Yaskawa INFORM job: ITEST.JBI

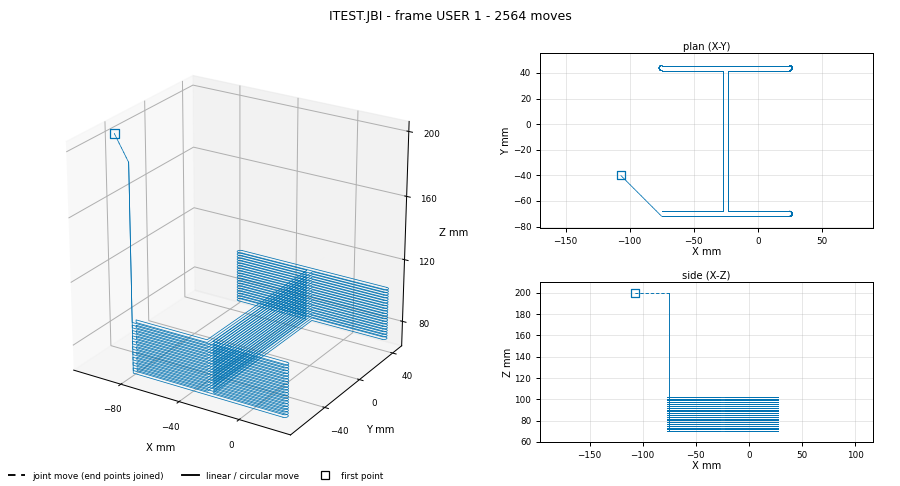
[picture p0: tool path of ITEST.JBI in frame USER 1, 2564 of 2624 moves have a stored position in this frame; points joined in program order, loops and branches not executed]
/JOB
//NAME ITEST
//POS
///NPOS 2624,0,0,0,0,0
///USER 1
///TOOL 1
///POSTYPE USER
///RECTAN
///RCONF 1,0,0,0,0,0,0,0,0,0,0,0,0,0,0,0,0,0,0,0,0,0,0,0
C00000=-107.000,-40.000,200.000,0.0000,0.0000,-150.0000
C00001=-75.000,-72.000,200.000,0.0000,0.0000,-150.0000
C00002=-75.000,-72.000,70.000,0.0000,0.0000,-150.0000
C00003=-70.000,-72.000,70.000,0.0000,0.0000,-150.0000
C00004=-65.000,-72.000,70.000,0.0000,0.0000,-150.0000
C00005=-60.000,-72.000,70.000,0.0000,0.0000,-150.0000
C00006=-55.000,-72.000,70.000,0.0000,0.0000,-150.0000
C00007=-50.000,-72.000,70.000,0.0000,0.0000,-150.0000
C00008=-45.000,-72.000,70.000,0.0000,0.0000,-150.0000
C00009=-40.000,-72.000,70.000,0.0000,0.0000,-150.0000
C00010=-35.000,-72.000,70.000,0.0000,0.0000,-150.0000
C00011=-30.000,-72.000,70.000,0.0000,0.0000,-150.0000
C00012=-25.000,-72.000,70.000,0.0000,0.0000,-150.0000
C00013=-20.000,-72.000,70.000,0.0000,0.0000,-150.0000
C00014=-15.000,-72.000,70.000,0.0000,0.0000,-150.0000
C00015=-10.000,-72.000,70.000,0.0000,0.0000,-150.0000
C00016=-5.000,-72.000,70.000,0.0000,0.0000,-150.0000
C00017=0.000,-72.000,70.000,0.0000,0.0000,-150.0000
C00018=5.000,-72.000,70.000,0.0000,0.0000,-150.0000
C00019=10.000,-72.000,70.000,0.0000,0.0000,-150.0000
C00020=15.000,-72.000,70.000,0.0000,0.0000,-150.0000
C00021=20.000,-72.000,70.000,0.0000,0.0000,-150.0000
C00022=25.000,-72.000,70.000,0.0000,0.0000,-150.0000
C00023=26.950,-70.050,70.000,0.0000,0.0000,-150.0000
C00024=25.000,-68.100,70.000,0.0000,0.0000,-150.0000
C00025=20.195,-68.100,70.000,0.0000,0.0000,-150.0000
C00026=15.390,-68.100,70.000,0.0000,0.0000,-150.0000
C00027=10.585,-68.100,70.000,0.0000,0.0000,-150.0000
C00028=5.780,-68.100,70.000,0.0000,0.0000,-150.0000
C00029=0.975,-68.100,70.000,0.0000,0.0000,-150.0000
C00030=-3.830,-68.100,70.000,0.0000,0.0000,-150.0000
C00031=-8.635,-68.100,70.000,0.0000,0.0000,-150.0000
C00032=-13.440,-68.100,70.000,0.0000,0.0000,-150.0000
C00033=-18.245,-68.100,70.000,0.0000,0.0000,-150.0000
C00034=-23.050,-68.100,70.000,0.0000,0.0000,-150.0000
C00035=-23.050,-63.100,70.000,0.0000,0.0000,-150.0000
C00036=-23.050,-58.100,70.000,0.0000,0.0000,-150.0000
C00037=-23.050,-53.100,70.000,0.0000,0.0000,-150.0000
C00038=-23.050,-48.100,70.000,0.0000,0.0000,-150.0000
C00039=-23.050,-43.100,70.000,0.0000,0.0000,-150.0000
C00040=-23.050,-38.100,70.000,0.0000,0.0000,-150.0000
C00041=-23.050,-33.100,70.000,0.0000,0.0000,-150.0000
C00042=-23.050,-28.100,70.000,0.0000,0.0000,-150.0000
C00043=-23.050,-23.100,70.000,0.0000,0.0000,-150.0000
C00044=-23.050,-18.100,70.000,0.0000,0.0000,-150.0000
C00045=-23.050,-13.100,70.000,0.0000,0.0000,-150.0000
C00046=-23.050,-8.100,70.000,0.0000,0.0000,-150.0000
C00047=-23.050,-3.100,70.000,0.0000,0.0000,-150.0000
C00048=-23.050,1.900,70.000,0.0000,0.0000,-150.0000
C00049=-23.050,6.900,70.000,0.0000,0.0000,-150.0000
C00050=-23.050,11.900,70.000,0.0000,0.0000,-150.0000
C00051=-23.050,16.900,70.000,0.0000,0.0000,-150.0000
C00052=-23.050,21.900,70.000,0.0000,0.0000,-150.0000
C00053=-23.050,26.900,70.000,0.0000,0.0000,-150.0000
C00054=-23.050,31.900,70.000,0.0000,0.0000,-150.0000
C00055=-23.050,36.900,70.000,0.0000,0.0000,-150.0000
C00056=-23.050,41.900,70.000,0.0000,0.0000,-150.0000
C00057=-18.267,41.900,70.000,0.0000,0.0000,-150.0000
C00058=-13.483,41.900,70.000,0.0000,0.0000,-150.0000
C00059=-8.700,41.900,70.000,0.0000,0.0000,-150.0000
C00060=-3.917,41.900,70.000,0.0000,0.0000,-150.0000
C00061=0.867,41.900,70.000,0.0000,0.0000,-150.0000
C00062=5.650,41.900,70.000,0.0000,0.0000,-150.0000
C00063=10.433,41.900,70.000,0.0000,0.0000,-150.0000
C00064=15.217,41.900,70.000,0.0000,0.0000,-150.0000
C00065=20.000,41.900,70.000,0.0000,0.0000,-150.0000
C00066=25.000,41.900,70.000,0.0000,0.0000,-150.0000
C00067=26.950,43.850,70.000,0.0000,0.0000,-150.0000
C00068=25.000,45.800,70.000,0.0000,0.0000,-150.0000
C00069=20.000,45.800,70.000,0.0000,0.0000,-150.0000
C00070=15.000,45.800,70.000,0.0000,0.0000,-150.0000
C00071=10.000,45.800,70.000,0.0000,0.0000,-150.0000
C00072=5.000,45.800,70.000,0.0000,0.0000,-150.0000
C00073=0.000,45.800,70.000,0.0000,0.0000,-150.0000
C00074=-5.000,45.800,70.000,0.0000,0.0000,-150.0000
C00075=-10.000,45.800,70.000,0.0000,0.0000,-150.0000
C00076=-15.000,45.800,70.000,0.0000,0.0000,-150.0000
C00077=-20.000,45.800,70.000,0.0000,0.0000,-150.0000
C00078=-25.000,45.800,70.000,0.0000,0.0000,-150.0000
C00079=-30.000,45.800,70.000,0.0000,0.0000,-150.0000
C00080=-35.000,45.800,70.000,0.0000,0.0000,-150.0000
C00081=-40.000,45.800,70.000,0.0000,0.0000,-150.0000
C00082=-45.000,45.800,70.000,0.0000,0.0000,-150.0000
C00083=-50.000,45.800,70.000,0.0000,0.0000,-150.0000
C00084=-55.000,45.800,70.000,0.0000,0.0000,-150.0000
C00085=-60.000,45.800,70.000,0.0000,0.0000,-150.0000
C00086=-65.000,45.800,70.000,0.0000,0.0000,-150.0000
C00087=-70.000,45.800,70.000,0.0000,0.0000,-150.0000
C00088=-75.000,45.800,70.000,0.0000,0.0000,-150.0000
C00089=-76.950,43.850,70.000,0.0000,0.0000,-150.0000
C00090=-75.000,41.900,70.000,0.0000,0.0000,-150.0000
C00091=-70.195,41.900,70.000,0.0000,0.0000,-150.0000
C00092=-65.390,41.900,70.000,0.0000,0.0000,-150.0000
C00093=-60.585,41.900,70.000,0.0000,0.0000,-150.0000
C00094=-55.780,41.900,70.000,0.0000,0.0000,-150.0000
C00095=-50.975,41.900,70.000,0.0000,0.0000,-150.0000
C00096=-46.170,41.900,70.000,0.0000,0.0000,-150.0000
C00097=-41.365,41.900,70.000,0.0000,0.0000,-150.0000
C00098=-36.560,41.900,70.000,0.0000,0.0000,-150.0000
C00099=-31.755,41.900,70.000,0.0000,0.0000,-150.0000
C00100=-26.950,41.900,70.000,0.0000,0.0000,-150.0000
C00101=-26.950,36.900,70.000,0.0000,0.0000,-150.0000
C00102=-26.950,31.900,70.000,0.0000,0.0000,-150.0000
C00103=-26.950,26.900,70.000,0.0000,0.0000,-150.0000
C00104=-26.950,21.900,70.000,0.0000,0.0000,-150.0000
C00105=-26.950,16.900,70.000,0.0000,0.0000,-150.0000
C00106=-26.950,11.900,70.000,0.0000,0.0000,-150.0000
C00107=-26.950,6.900,70.000,0.0000,0.0000,-150.0000
C00108=-26.950,1.900,70.000,0.0000,0.0000,-150.0000
C00109=-26.950,-3.100,70.000,0.0000,0.0000,-150.0000
C00110=-26.950,-8.100,70.000,0.0000,0.0000,-150.0000
C00111=-26.950,-13.100,70.000,0.0000,0.0000,-150.0000
C00112=-26.950,-18.100,70.000,0.0000,0.0000,-150.0000
C00113=-26.950,-23.100,70.000,0.0000,0.0000,-150.0000
C00114=-26.950,-28.100,70.000,0.0000,0.0000,-150.0000
C00115=-26.950,-33.100,70.000,0.0000,0.0000,-150.0000
C00116=-26.950,-38.100,70.000,0.0000,0.0000,-150.0000
C00117=-26.950,-43.100,70.000,0.0000,0.0000,-150.0000
C00118=-26.950,-48.100,70.000,0.0000,0.0000,-150.0000
C00119=-26.950,-53.100,70.000,0.0000,0.0000,-150.0000
C00120=-26.950,-58.100,70.000,0.0000,0.0000,-150.0000
C00121=-26.950,-63.100,70.000,0.0000,0.0000,-150.0000
C00122=-26.950,-68.100,70.000,0.0000,0.0000,-150.0000
C00123=-31.755,-68.100,70.000,0.0000,0.0000,-150.0000
C00124=-36.560,-68.100,70.000,0.0000,0.0000,-150.0000
C00125=-41.365,-68.100,70.000,0.0000,0.0000,-150.0000
C00126=-46.170,-68.100,70.000,0.0000,0.0000,-150.0000
C00127=-50.975,-68.100,70.000,0.0000,0.0000,-150.0000
C00128=-55.780,-68.100,70.000,0.0000,0.0000,-150.0000
C00129=-60.585,-68.100,70.000,0.0000,0.0000,-150.0000
C00130=-65.390,-68.100,70.000,0.0000,0.0000,-150.0000
C00131=-70.195,-68.100,70.000,0.0000,0.0000,-150.0000
C00132=-75.000,-68.100,70.000,0.0000,0.0000,-150.0000
C00133=-75.000,-68.100,71.700,0.0000,0.0000,-150.0000
C00134=-70.195,-68.100,71.700,0.0000,0.0000,-150.0000
C00135=-65.390,-68.100,71.700,0.0000,0.0000,-150.0000
C00136=-60.585,-68.100,71.700,0.0000,0.0000,-150.0000
C00137=-55.780,-68.100,71.700,0.0000,0.0000,-150.0000
C00138=-50.975,-68.100,71.700,0.0000,0.0000,-150.0000
C00139=-46.170,-68.100,71.700,0.0000,0.0000,-150.0000
C00140=-41.365,-68.100,71.700,0.0000,0.0000,-150.0000
C00141=-36.560,-68.100,71.700,0.0000,0.0000,-150.0000
C00142=-31.755,-68.100,71.700,0.0000,0.0000,-150.0000
C00143=-26.950,-68.100,71.700,0.0000,0.0000,-150.0000
C00144=-26.950,-63.100,71.700,0.0000,0.0000,-150.0000
C00145=-26.950,-58.100,71.700,0.0000,0.0000,-150.0000
C00146=-26.950,-53.100,71.700,0.0000,0.0000,-150.0000
C00147=-26.950,-48.100,71.700,0.0000,0.0000,-150.0000
C00148=-26.950,-43.100,71.700,0.0000,0.0000,-150.0000
C00149=-26.950,-38.100,71.700,0.0000,0.0000,-150.0000
C00150=-26.950,-33.100,71.700,0.0000,0.0000,-150.0000
C00151=-26.950,-28.100,71.700,0.0000,0.0000,-150.0000
C00152=-26.950,-23.100,71.700,0.0000,0.0000,-150.0000
C00153=-26.950,-18.100,71.700,0.0000,0.0000,-150.0000
C00154=-26.950,-13.100,71.700,0.0000,0.0000,-150.0000
C00155=-26.950,-8.100,71.700,0.0000,0.0000,-150.0000
C00156=-26.950,-3.100,71.700,0.0000,0.0000,-150.0000
C00157=-26.950,1.900,71.700,0.0000,0.0000,-150.0000
C00158=-26.950,6.900,71.700,0.0000,0.0000,-150.0000
C00159=-26.950,11.900,71.700,0.0000,0.0000,-150.0000
C00160=-26.950,16.900,71.700,0.0000,0.0000,-150.0000
C00161=-26.950,21.900,71.700,0.0000,0.0000,-150.0000
C00162=-26.950,26.900,71.700,0.0000,0.0000,-150.0000
C00163=-26.950,31.900,71.700,0.0000,0.0000,-150.0000
C00164=-26.950,36.900,71.700,0.0000,0.0000,-150.0000
C00165=-26.950,41.900,71.700,0.0000,0.0000,-150.0000
C00166=-31.733,41.900,71.700,0.0000,0.0000,-150.0000
C00167=-36.517,41.900,71.700,0.0000,0.0000,-150.0000
C00168=-41.300,41.900,71.700,0.0000,0.0000,-150.0000
C00169=-46.083,41.900,71.700,0.0000,0.0000,-150.0000
C00170=-50.867,41.900,71.700,0.0000,0.0000,-150.0000
C00171=-55.650,41.900,71.700,0.0000,0.0000,-150.0000
C00172=-60.433,41.900,71.700,0.0000,0.0000,-150.0000
C00173=-65.217,41.900,71.700,0.0000,0.0000,-150.0000
C00174=-70.000,41.900,71.700,0.0000,0.0000,-150.0000
C00175=-75.000,41.900,71.700,0.0000,0.0000,-150.0000
C00176=-76.950,43.850,71.700,0.0000,0.0000,-150.0000
C00177=-75.000,45.800,71.700,0.0000,0.0000,-150.0000
C00178=-70.000,45.800,71.700,0.0000,0.0000,-150.0000
C00179=-65.000,45.800,71.700,0.0000,0.0000,-150.0000
C00180=-60.000,45.800,71.700,0.0000,0.0000,-150.0000
C00181=-55.000,45.800,71.700,0.0000,0.0000,-150.0000
C00182=-50.000,45.800,71.700,0.0000,0.0000,-150.0000
C00183=-45.000,45.800,71.700,0.0000,0.0000,-150.0000
C00184=-40.000,45.800,71.700,0.0000,0.0000,-150.0000
C00185=-35.000,45.800,71.700,0.0000,0.0000,-150.0000
C00186=-30.000,45.800,71.700,0.0000,0.0000,-150.0000
C00187=-25.000,45.800,71.700,0.0000,0.0000,-150.0000
C00188=-20.000,45.800,71.700,0.0000,0.0000,-150.0000
C00189=-15.000,45.800,71.700,0.0000,0.0000,-150.0000
C00190=-10.000,45.800,71.700,0.0000,0.0000,-150.0000
C00191=-5.000,45.800,71.700,0.0000,0.0000,-150.0000
C00192=0.000,45.800,71.700,0.0000,0.0000,-150.0000
C00193=5.000,45.800,71.700,0.0000,0.0000,-150.0000
C00194=10.000,45.800,71.700,0.0000,0.0000,-150.0000
C00195=15.000,45.800,71.700,0.0000,0.0000,-150.0000
C00196=20.000,45.800,71.700,0.0000,0.0000,-150.0000
C00197=25.000,45.800,71.700,0.0000,0.0000,-150.0000
C00198=26.950,43.850,71.700,0.0000,0.0000,-150.0000
C00199=25.000,41.900,71.700,0.0000,0.0000,-150.0000
C00200=20.195,41.900,71.700,0.0000,0.0000,-150.0000
C00201=15.390,41.900,71.700,0.0000,0.0000,-150.0000
C00202=10.585,41.900,71.700,0.0000,0.0000,-150.0000
C00203=5.780,41.900,71.700,0.0000,0.0000,-150.0000
C00204=0.975,41.900,71.700,0.0000,0.0000,-150.0000
C00205=-3.830,41.900,71.700,0.0000,0.0000,-150.0000
C00206=-8.635,41.900,71.700,0.0000,0.0000,-150.0000
C00207=-13.440,41.900,71.700,0.0000,0.0000,-150.0000
C00208=-18.245,41.900,71.700,0.0000,0.0000,-150.0000
C00209=-23.050,41.900,71.700,0.0000,0.0000,-150.0000
C00210=-23.050,36.900,71.700,0.0000,0.0000,-150.0000
C00211=-23.050,31.900,71.700,0.0000,0.0000,-150.0000
C00212=-23.050,26.900,71.700,0.0000,0.0000,-150.0000
C00213=-23.050,21.900,71.700,0.0000,0.0000,-150.0000
C00214=-23.050,16.900,71.700,0.0000,0.0000,-150.0000
C00215=-23.050,11.900,71.700,0.0000,0.0000,-150.0000
C00216=-23.050,6.900,71.700,0.0000,0.0000,-150.0000
C00217=-23.050,1.900,71.700,0.0000,0.0000,-150.0000
C00218=-23.050,-3.100,71.700,0.0000,0.0000,-150.0000
C00219=-23.050,-8.100,71.700,0.0000,0.0000,-150.0000
C00220=-23.050,-13.100,71.700,0.0000,0.0000,-150.0000
C00221=-23.050,-18.100,71.700,0.0000,0.0000,-150.0000
C00222=-23.050,-23.100,71.700,0.0000,0.0000,-150.0000
C00223=-23.050,-28.100,71.700,0.0000,0.0000,-150.0000
C00224=-23.050,-33.100,71.700,0.0000,0.0000,-150.0000
C00225=-23.050,-38.100,71.700,0.0000,0.0000,-150.0000
C00226=-23.050,-43.100,71.700,0.0000,0.0000,-150.0000
C00227=-23.050,-48.100,71.700,0.0000,0.0000,-150.0000
C00228=-23.050,-53.100,71.700,0.0000,0.0000,-150.0000
C00229=-23.050,-58.100,71.700,0.0000,0.0000,-150.0000
C00230=-23.050,-63.100,71.700,0.0000,0.0000,-150.0000
C00231=-23.050,-68.100,71.700,0.0000,0.0000,-150.0000
C00232=-18.267,-68.100,71.700,0.0000,0.0000,-150.0000
C00233=-13.483,-68.100,71.700,0.0000,0.0000,-150.0000
C00234=-8.700,-68.100,71.700,0.0000,0.0000,-150.0000
C00235=-3.917,-68.100,71.700,0.0000,0.0000,-150.0000
C00236=0.867,-68.100,71.700,0.0000,0.0000,-150.0000
C00237=5.650,-68.100,71.700,0.0000,0.0000,-150.0000
C00238=10.433,-68.100,71.700,0.0000,0.0000,-150.0000
C00239=15.217,-68.100,71.700,0.0000,0.0000,-150.0000
C00240=20.000,-68.100,71.700,0.0000,0.0000,-150.0000
C00241=25.000,-68.100,71.700,0.0000,0.0000,-150.0000
C00242=26.950,-70.050,71.700,0.0000,0.0000,-150.0000
C00243=25.000,-72.000,71.700,0.0000,0.0000,-150.0000
C00244=20.000,-72.000,71.700,0.0000,0.0000,-150.0000
C00245=15.000,-72.000,71.700,0.0000,0.0000,-150.0000
C00246=10.000,-72.000,71.700,0.0000,0.0000,-150.0000
C00247=5.000,-72.000,71.700,0.0000,0.0000,-150.0000
C00248=0.000,-72.000,71.700,0.0000,0.0000,-150.0000
C00249=-5.000,-72.000,71.700,0.0000,0.0000,-150.0000
C00250=-10.000,-72.000,71.700,0.0000,0.0000,-150.0000
C00251=-15.000,-72.000,71.700,0.0000,0.0000,-150.0000
C00252=-20.000,-72.000,71.700,0.0000,0.0000,-150.0000
C00253=-25.000,-72.000,71.700,0.0000,0.0000,-150.0000
C00254=-30.000,-72.000,71.700,0.0000,0.0000,-150.0000
C00255=-35.000,-72.000,71.700,0.0000,0.0000,-150.0000
C00256=-40.000,-72.000,71.700,0.0000,0.0000,-150.0000
C00257=-45.000,-72.000,71.700,0.0000,0.0000,-150.0000
C00258=-50.000,-72.000,71.700,0.0000,0.0000,-150.0000
C00259=-55.000,-72.000,71.700,0.0000,0.0000,-150.0000
C00260=-60.000,-72.000,71.700,0.0000,0.0000,-150.0000
C00261=-65.000,-72.000,71.700,0.0000,0.0000,-150.0000
C00262=-70.000,-72.000,71.700,0.0000,0.0000,-150.0000
C00263=-75.000,-72.000,71.700,0.0000,0.0000,-150.0000
C00264=-75.000,-72.000,73.400,0.0000,0.0000,-150.0000
C00265=-70.000,-72.000,73.400,0.0000,0.0000,-150.0000
C00266=-65.000,-72.000,73.400,0.0000,0.0000,-150.0000
C00267=-60.000,-72.000,73.400,0.0000,0.0000,-150.0000
C00268=-55.000,-72.000,73.400,0.0000,0.0000,-150.0000
C00269=-50.000,-72.000,73.400,0.0000,0.0000,-150.0000
C00270=-45.000,-72.000,73.400,0.0000,0.0000,-150.0000
C00271=-40.000,-72.000,73.400,0.0000,0.0000,-150.0000
C00272=-35.000,-72.000,73.400,0.0000,0.0000,-150.0000
C00273=-30.000,-72.000,73.400,0.0000,0.0000,-150.0000
C00274=-25.000,-72.000,73.400,0.0000,0.0000,-150.0000
C00275=-20.000,-72.000,73.400,0.0000,0.0000,-150.0000
C00276=-15.000,-72.000,73.400,0.0000,0.0000,-150.0000
C00277=-10.000,-72.000,73.400,0.0000,0.0000,-150.0000
C00278=-5.000,-72.000,73.400,0.0000,0.0000,-150.0000
C00279=0.000,-72.000,73.400,0.0000,0.0000,-150.0000
C00280=5.000,-72.000,73.400,0.0000,0.0000,-150.0000
C00281=10.000,-72.000,73.400,0.0000,0.0000,-150.0000
C00282=15.000,-72.000,73.400,0.0000,0.0000,-150.0000
C00283=20.000,-72.000,73.400,0.0000,0.0000,-150.0000
C00284=25.000,-72.000,73.400,0.0000,0.0000,-150.0000
C00285=26.950,-70.050,73.400,0.0000,0.0000,-150.0000
C00286=25.000,-68.100,73.400,0.0000,0.0000,-150.0000
C00287=20.195,-68.100,73.400,0.0000,0.0000,-150.0000
C00288=15.390,-68.100,73.400,0.0000,0.0000,-150.0000
C00289=10.585,-68.100,73.400,0.0000,0.0000,-150.0000
C00290=5.780,-68.100,73.400,0.0000,0.0000,-150.0000
C00291=0.975,-68.100,73.400,0.0000,0.0000,-150.0000
C00292=-3.830,-68.100,73.400,0.0000,0.0000,-150.0000
C00293=-8.635,-68.100,73.400,0.0000,0.0000,-150.0000
C00294=-13.440,-68.100,73.400,0.0000,0.0000,-150.0000
C00295=-18.245,-68.100,73.400,0.0000,0.0000,-150.0000
C00296=-23.050,-68.100,73.400,0.0000,0.0000,-150.0000
C00297=-23.050,-63.100,73.400,0.0000,0.0000,-150.0000
C00298=-23.050,-58.100,73.400,0.0000,0.0000,-150.0000
C00299=-23.050,-53.100,73.400,0.0000,0.0000,-150.0000
C00300=-23.050,-48.100,73.400,0.0000,0.0000,-150.0000
C00301=-23.050,-43.100,73.400,0.0000,0.0000,-150.0000
C00302=-23.050,-38.100,73.400,0.0000,0.0000,-150.0000
C00303=-23.050,-33.100,73.400,0.0000,0.0000,-150.0000
C00304=-23.050,-28.100,73.400,0.0000,0.0000,-150.0000
C00305=-23.050,-23.100,73.400,0.0000,0.0000,-150.0000
C00306=-23.050,-18.100,73.400,0.0000,0.0000,-150.0000
C00307=-23.050,-13.100,73.400,0.0000,0.0000,-150.0000
C00308=-23.050,-8.100,73.400,0.0000,0.0000,-150.0000
C00309=-23.050,-3.100,73.400,0.0000,0.0000,-150.0000
C00310=-23.050,1.900,73.400,0.0000,0.0000,-150.0000
C00311=-23.050,6.900,73.400,0.0000,0.0000,-150.0000
C00312=-23.050,11.900,73.400,0.0000,0.0000,-150.0000
C00313=-23.050,16.900,73.400,0.0000,0.0000,-150.0000
C00314=-23.050,21.900,73.400,0.0000,0.0000,-150.0000
C00315=-23.050,26.900,73.400,0.0000,0.0000,-150.0000
C00316=-23.050,31.900,73.400,0.0000,0.0000,-150.0000
C00317=-23.050,36.900,73.400,0.0000,0.0000,-150.0000
C00318=-23.050,41.900,73.400,0.0000,0.0000,-150.0000
C00319=-18.267,41.900,73.400,0.0000,0.0000,-150.0000
C00320=-13.483,41.900,73.400,0.0000,0.0000,-150.0000
C00321=-8.700,41.900,73.400,0.0000,0.0000,-150.0000
C00322=-3.917,41.900,73.400,0.0000,0.0000,-150.0000
C00323=0.867,41.900,73.400,0.0000,0.0000,-150.0000
C00324=5.650,41.900,73.400,0.0000,0.0000,-150.0000
C00325=10.433,41.900,73.400,0.0000,0.0000,-150.0000
C00326=15.217,41.900,73.400,0.0000,0.0000,-150.0000
C00327=20.000,41.900,73.400,0.0000,0.0000,-150.0000
C00328=25.000,41.900,73.400,0.0000,0.0000,-150.0000
C00329=26.950,43.850,73.400,0.0000,0.0000,-150.0000
C00330=25.000,45.800,73.400,0.0000,0.0000,-150.0000
C00331=20.000,45.800,73.400,0.0000,0.0000,-150.0000
C00332=15.000,45.800,73.400,0.0000,0.0000,-150.0000
C00333=10.000,45.800,73.400,0.0000,0.0000,-150.0000
C00334=5.000,45.800,73.400,0.0000,0.0000,-150.0000
C00335=0.000,45.800,73.400,0.0000,0.0000,-150.0000
C00336=-5.000,45.800,73.400,0.0000,0.0000,-150.0000
C00337=-10.000,45.800,73.400,0.0000,0.0000,-150.0000
C00338=-15.000,45.800,73.400,0.0000,0.0000,-150.0000
C00339=-20.000,45.800,73.400,0.0000,0.0000,-150.0000
C00340=-25.000,45.800,73.400,0.0000,0.0000,-150.0000
C00341=-30.000,45.800,73.400,0.0000,0.0000,-150.0000
C00342=-35.000,45.800,73.400,0.0000,0.0000,-150.0000
C00343=-40.000,45.800,73.400,0.0000,0.0000,-150.0000
C00344=-45.000,45.800,73.400,0.0000,0.0000,-150.0000
C00345=-50.000,45.800,73.400,0.0000,0.0000,-150.0000
C00346=-55.000,45.800,73.400,0.0000,0.0000,-150.0000
C00347=-60.000,45.800,73.400,0.0000,0.0000,-150.0000
C00348=-65.000,45.800,73.400,0.0000,0.0000,-150.0000
C00349=-70.000,45.800,73.400,0.0000,0.0000,-150.0000
C00350=-75.000,45.800,73.400,0.0000,0.0000,-150.0000
C00351=-76.950,43.850,73.400,0.0000,0.0000,-150.0000
C00352=-75.000,41.900,73.400,0.0000,0.0000,-150.0000
C00353=-70.195,41.900,73.400,0.0000,0.0000,-150.0000
C00354=-65.390,41.900,73.400,0.0000,0.0000,-150.0000
C00355=-60.585,41.900,73.400,0.0000,0.0000,-150.0000
C00356=-55.780,41.900,73.400,0.0000,0.0000,-150.0000
C00357=-50.975,41.900,73.400,0.0000,0.0000,-150.0000
C00358=-46.170,41.900,73.400,0.0000,0.0000,-150.0000
C00359=-41.365,41.900,73.400,0.0000,0.0000,-150.0000
C00360=-36.560,41.900,73.400,0.0000,0.0000,-150.0000
C00361=-31.755,41.900,73.400,0.0000,0.0000,-150.0000
C00362=-26.950,41.900,73.400,0.0000,0.0000,-150.0000
C00363=-26.950,36.900,73.400,0.0000,0.0000,-150.0000
C00364=-26.950,31.900,73.400,0.0000,0.0000,-150.0000
C00365=-26.950,26.900,73.400,0.0000,0.0000,-150.0000
C00366=-26.950,21.900,73.400,0.0000,0.0000,-150.0000
C00367=-26.950,16.900,73.400,0.0000,0.0000,-150.0000
C00368=-26.950,11.900,73.400,0.0000,0.0000,-150.0000
C00369=-26.950,6.900,73.400,0.0000,0.0000,-150.0000
C00370=-26.950,1.900,73.400,0.0000,0.0000,-150.0000
C00371=-26.950,-3.100,73.400,0.0000,0.0000,-150.0000
C00372=-26.950,-8.100,73.400,0.0000,0.0000,-150.0000
C00373=-26.950,-13.100,73.400,0.0000,0.0000,-150.0000
C00374=-26.950,-18.100,73.400,0.0000,0.0000,-150.0000
C00375=-26.950,-23.100,73.400,0.0000,0.0000,-150.0000
C00376=-26.950,-28.100,73.400,0.0000,0.0000,-150.0000
C00377=-26.950,-33.100,73.400,0.0000,0.0000,-150.0000
C00378=-26.950,-38.100,73.400,0.0000,0.0000,-150.0000
C00379=-26.950,-43.100,73.400,0.0000,0.0000,-150.0000
C00380=-26.950,-48.100,73.400,0.0000,0.0000,-150.0000
C00381=-26.950,-53.100,73.400,0.0000,0.0000,-150.0000
C00382=-26.950,-58.100,73.400,0.0000,0.0000,-150.0000
C00383=-26.950,-63.100,73.400,0.0000,0.0000,-150.0000
C00384=-26.950,-68.100,73.400,0.0000,0.0000,-150.0000
C00385=-31.755,-68.100,73.400,0.0000,0.0000,-150.0000
C00386=-36.560,-68.100,73.400,0.0000,0.0000,-150.0000
C00387=-41.365,-68.100,73.400,0.0000,0.0000,-150.0000
C00388=-46.170,-68.100,73.400,0.0000,0.0000,-150.0000
C00389=-50.975,-68.100,73.400,0.0000,0.0000,-150.0000
C00390=-55.780,-68.100,73.400,0.0000,0.0000,-150.0000
C00391=-60.585,-68.100,73.400,0.0000,0.0000,-150.0000
C00392=-65.390,-68.100,73.400,0.0000,0.0000,-150.0000
C00393=-70.195,-68.100,73.400,0.0000,0.0000,-150.0000
C00394=-75.000,-68.100,73.400,0.0000,0.0000,-150.0000
C00395=-75.000,-68.100,75.100,0.0000,0.0000,-150.0000
C00396=-70.195,-68.100,75.100,0.0000,0.0000,-150.0000
C00397=-65.390,-68.100,75.100,0.0000,0.0000,-150.0000
C00398=-60.585,-68.100,75.100,0.0000,0.0000,-150.0000
C00399=-55.780,-68.100,75.100,0.0000,0.0000,-150.0000
C00400=-50.975,-68.100,75.100,0.0000,0.0000,-150.0000
C00401=-46.170,-68.100,75.100,0.0000,0.0000,-150.0000
C00402=-41.365,-68.100,75.100,0.0000,0.0000,-150.0000
C00403=-36.560,-68.100,75.100,0.0000,0.0000,-150.0000
C00404=-31.755,-68.100,75.100,0.0000,0.0000,-150.0000
C00405=-26.950,-68.100,75.100,0.0000,0.0000,-150.0000
C00406=-26.950,-63.100,75.100,0.0000,0.0000,-150.0000
C00407=-26.950,-58.100,75.100,0.0000,0.0000,-150.0000
C00408=-26.950,-53.100,75.100,0.0000,0.0000,-150.0000
C00409=-26.950,-48.100,75.100,0.0000,0.0000,-150.0000
C00410=-26.950,-43.100,75.100,0.0000,0.0000,-150.0000
C00411=-26.950,-38.100,75.100,0.0000,0.0000,-150.0000
C00412=-26.950,-33.100,75.100,0.0000,0.0000,-150.0000
C00413=-26.950,-28.100,75.100,0.0000,0.0000,-150.0000
C00414=-26.950,-23.100,75.100,0.0000,0.0000,-150.0000
C00415=-26.950,-18.100,75.100,0.0000,0.0000,-150.0000
C00416=-26.950,-13.100,75.100,0.0000,0.0000,-150.0000
C00417=-26.950,-8.100,75.100,0.0000,0.0000,-150.0000
C00418=-26.950,-3.100,75.100,0.0000,0.0000,-150.0000
C00419=-26.950,1.900,75.100,0.0000,0.0000,-150.0000
C00420=-26.950,6.900,75.100,0.0000,0.0000,-150.0000
C00421=-26.950,11.900,75.100,0.0000,0.0000,-150.0000
C00422=-26.950,16.900,75.100,0.0000,0.0000,-150.0000
C00423=-26.950,21.900,75.100,0.0000,0.0000,-150.0000
C00424=-26.950,26.900,75.100,0.0000,0.0000,-150.0000
C00425=-26.950,31.900,75.100,0.0000,0.0000,-150.0000
C00426=-26.950,36.900,75.100,0.0000,0.0000,-150.0000
C00427=-26.950,41.900,75.100,0.0000,0.0000,-150.0000
C00428=-31.733,41.900,75.100,0.0000,0.0000,-150.0000
C00429=-36.517,41.900,75.100,0.0000,0.0000,-150.0000
C00430=-41.300,41.900,75.100,0.0000,0.0000,-150.0000
C00431=-46.083,41.900,75.100,0.0000,0.0000,-150.0000
C00432=-50.867,41.900,75.100,0.0000,0.0000,-150.0000
C00433=-55.650,41.900,75.100,0.0000,0.0000,-150.0000
C00434=-60.433,41.900,75.100,0.0000,0.0000,-150.0000
C00435=-65.217,41.900,75.100,0.0000,0.0000,-150.0000
C00436=-70.000,41.900,75.100,0.0000,0.0000,-150.0000
C00437=-75.000,41.900,75.100,0.0000,0.0000,-150.0000
C00438=-76.950,43.850,75.100,0.0000,0.0000,-150.0000
C00439=-75.000,45.800,75.100,0.0000,0.0000,-150.0000
C00440=-70.000,45.800,75.100,0.0000,0.0000,-150.0000
C00441=-65.000,45.800,75.100,0.0000,0.0000,-150.0000
C00442=-60.000,45.800,75.100,0.0000,0.0000,-150.0000
C00443=-55.000,45.800,75.100,0.0000,0.0000,-150.0000
C00444=-50.000,45.800,75.100,0.0000,0.0000,-150.0000
C00445=-45.000,45.800,75.100,0.0000,0.0000,-150.0000
C00446=-40.000,45.800,75.100,0.0000,0.0000,-150.0000
C00447=-35.000,45.800,75.100,0.0000,0.0000,-150.0000
C00448=-30.000,45.800,75.100,0.0000,0.0000,-150.0000
C00449=-25.000,45.800,75.100,0.0000,0.0000,-150.0000
C00450=-20.000,45.800,75.100,0.0000,0.0000,-150.0000
C00451=-15.000,45.800,75.100,0.0000,0.0000,-150.0000
C00452=-10.000,45.800,75.100,0.0000,0.0000,-150.0000
C00453=-5.000,45.800,75.100,0.0000,0.0000,-150.0000
C00454=0.000,45.800,75.100,0.0000,0.0000,-150.0000
C00455=5.000,45.800,75.100,0.0000,0.0000,-150.0000
C00456=10.000,45.800,75.100,0.0000,0.0000,-150.0000
C00457=15.000,45.800,75.100,0.0000,0.0000,-150.0000
C00458=20.000,45.800,75.100,0.0000,0.0000,-150.0000
C00459=25.000,45.800,75.100,0.0000,0.0000,-150.0000
C00460=26.950,43.850,75.100,0.0000,0.0000,-150.0000
C00461=25.000,41.900,75.100,0.0000,0.0000,-150.0000
C00462=20.195,41.900,75.100,0.0000,0.0000,-150.0000
C00463=15.390,41.900,75.100,0.0000,0.0000,-150.0000
C00464=10.585,41.900,75.100,0.0000,0.0000,-150.0000
C00465=5.780,41.900,75.100,0.0000,0.0000,-150.0000
C00466=0.975,41.900,75.100,0.0000,0.0000,-150.0000
C00467=-3.830,41.900,75.100,0.0000,0.0000,-150.0000
C00468=-8.635,41.900,75.100,0.0000,0.0000,-150.0000
C00469=-13.440,41.900,75.100,0.0000,0.0000,-150.0000
C00470=-18.245,41.900,75.100,0.0000,0.0000,-150.0000
C00471=-23.050,41.900,75.100,0.0000,0.0000,-150.0000
C00472=-23.050,36.900,75.100,0.0000,0.0000,-150.0000
C00473=-23.050,31.900,75.100,0.0000,0.0000,-150.0000
C00474=-23.050,26.900,75.100,0.0000,0.0000,-150.0000
C00475=-23.050,21.900,75.100,0.0000,0.0000,-150.0000
C00476=-23.050,16.900,75.100,0.0000,0.0000,-150.0000
C00477=-23.050,11.900,75.100,0.0000,0.0000,-150.0000
C00478=-23.050,6.900,75.100,0.0000,0.0000,-150.0000
C00479=-23.050,1.900,75.100,0.0000,0.0000,-150.0000
C00480=-23.050,-3.100,75.100,0.0000,0.0000,-150.0000
C00481=-23.050,-8.100,75.100,0.0000,0.0000,-150.0000
C00482=-23.050,-13.100,75.100,0.0000,0.0000,-150.0000
C00483=-23.050,-18.100,75.100,0.0000,0.0000,-150.0000
C00484=-23.050,-23.100,75.100,0.0000,0.0000,-150.0000
C00485=-23.050,-28.100,75.100,0.0000,0.0000,-150.0000
C00486=-23.050,-33.100,75.100,0.0000,0.0000,-150.0000
C00487=-23.050,-38.100,75.100,0.0000,0.0000,-150.0000
C00488=-23.050,-43.100,75.100,0.0000,0.0000,-150.0000
C00489=-23.050,-48.100,75.100,0.0000,0.0000,-150.0000
C00490=-23.050,-53.100,75.100,0.0000,0.0000,-150.0000
C00491=-23.050,-58.100,75.100,0.0000,0.0000,-150.0000
C00492=-23.050,-63.100,75.100,0.0000,0.0000,-150.0000
C00493=-23.050,-68.100,75.100,0.0000,0.0000,-150.0000
C00494=-18.267,-68.100,75.100,0.0000,0.0000,-150.0000
C00495=-13.483,-68.100,75.100,0.0000,0.0000,-150.0000
C00496=-8.700,-68.100,75.100,0.0000,0.0000,-150.0000
C00497=-3.917,-68.100,75.100,0.0000,0.0000,-150.0000
C00498=0.867,-68.100,75.100,0.0000,0.0000,-150.0000
C00499=5.650,-68.100,75.100,0.0000,0.0000,-150.0000
C00500=10.433,-68.100,75.100,0.0000,0.0000,-150.0000
C00501=15.217,-68.100,75.100,0.0000,0.0000,-150.0000
C00502=20.000,-68.100,75.100,0.0000,0.0000,-150.0000
C00503=25.000,-68.100,75.100,0.0000,0.0000,-150.0000
C00504=26.950,-70.050,75.100,0.0000,0.0000,-150.0000
C00505=25.000,-72.000,75.100,0.0000,0.0000,-150.0000
C00506=20.000,-72.000,75.100,0.0000,0.0000,-150.0000
C00507=15.000,-72.000,75.100,0.0000,0.0000,-150.0000
C00508=10.000,-72.000,75.100,0.0000,0.0000,-150.0000
C00509=5.000,-72.000,75.100,0.0000,0.0000,-150.0000
C00510=0.000,-72.000,75.100,0.0000,0.0000,-150.0000
C00511=-5.000,-72.000,75.100,0.0000,0.0000,-150.0000
C00512=-10.000,-72.000,75.100,0.0000,0.0000,-150.0000
C00513=-15.000,-72.000,75.100,0.0000,0.0000,-150.0000
C00514=-20.000,-72.000,75.100,0.0000,0.0000,-150.0000
C00515=-25.000,-72.000,75.100,0.0000,0.0000,-150.0000
C00516=-30.000,-72.000,75.100,0.0000,0.0000,-150.0000
C00517=-35.000,-72.000,75.100,0.0000,0.0000,-150.0000
C00518=-40.000,-72.000,75.100,0.0000,0.0000,-150.0000
C00519=-45.000,-72.000,75.100,0.0000,0.0000,-150.0000
C00520=-50.000,-72.000,75.100,0.0000,0.0000,-150.0000
C00521=-55.000,-72.000,75.100,0.0000,0.0000,-150.0000
C00522=-60.000,-72.000,75.100,0.0000,0.0000,-150.0000
C00523=-65.000,-72.000,75.100,0.0000,0.0000,-150.0000
C00524=-70.000,-72.000,75.100,0.0000,0.0000,-150.0000
C00525=-75.000,-72.000,75.100,0.0000,0.0000,-150.0000
C00526=-75.000,-72.000,76.800,0.0000,0.0000,-150.0000
C00527=-70.000,-72.000,76.800,0.0000,0.0000,-150.0000
C00528=-65.000,-72.000,76.800,0.0000,0.0000,-150.0000
C00529=-60.000,-72.000,76.800,0.0000,0.0000,-150.0000
C00530=-55.000,-72.000,76.800,0.0000,0.0000,-150.0000
C00531=-50.000,-72.000,76.800,0.0000,0.0000,-150.0000
C00532=-45.000,-72.000,76.800,0.0000,0.0000,-150.0000
C00533=-40.000,-72.000,76.800,0.0000,0.0000,-150.0000
C00534=-35.000,-72.000,76.800,0.0000,0.0000,-150.0000
C00535=-30.000,-72.000,76.800,0.0000,0.0000,-150.0000
C00536=-25.000,-72.000,76.800,0.0000,0.0000,-150.0000
C00537=-20.000,-72.000,76.800,0.0000,0.0000,-150.0000
C00538=-15.000,-72.000,76.800,0.0000,0.0000,-150.0000
C00539=-10.000,-72.000,76.800,0.0000,0.0000,-150.0000
C00540=-5.000,-72.000,76.800,0.0000,0.0000,-150.0000
C00541=0.000,-72.000,76.800,0.0000,0.0000,-150.0000
C00542=5.000,-72.000,76.800,0.0000,0.0000,-150.0000
C00543=10.000,-72.000,76.800,0.0000,0.0000,-150.0000
C00544=15.000,-72.000,76.800,0.0000,0.0000,-150.0000
C00545=20.000,-72.000,76.800,0.0000,0.0000,-150.0000
C00546=25.000,-72.000,76.800,0.0000,0.0000,-150.0000
C00547=26.950,-70.050,76.800,0.0000,0.0000,-150.0000
C00548=25.000,-68.100,76.800,0.0000,0.0000,-150.0000
C00549=20.195,-68.100,76.800,0.0000,0.0000,-150.0000
C00550=15.390,-68.100,76.800,0.0000,0.0000,-150.0000
C00551=10.585,-68.100,76.800,0.0000,0.0000,-150.0000
C00552=5.780,-68.100,76.800,0.0000,0.0000,-150.0000
C00553=0.975,-68.100,76.800,0.0000,0.0000,-150.0000
C00554=-3.830,-68.100,76.800,0.0000,0.0000,-150.0000
C00555=-8.635,-68.100,76.800,0.0000,0.0000,-150.0000
C00556=-13.440,-68.100,76.800,0.0000,0.0000,-150.0000
C00557=-18.245,-68.100,76.800,0.0000,0.0000,-150.0000
C00558=-23.050,-68.100,76.800,0.0000,0.0000,-150.0000
C00559=-23.050,-63.100,76.800,0.0000,0.0000,-150.0000
C00560=-23.050,-58.100,76.800,0.0000,0.0000,-150.0000
C00561=-23.050,-53.100,76.800,0.0000,0.0000,-150.0000
C00562=-23.050,-48.100,76.800,0.0000,0.0000,-150.0000
C00563=-23.050,-43.100,76.800,0.0000,0.0000,-150.0000
C00564=-23.050,-38.100,76.800,0.0000,0.0000,-150.0000
C00565=-23.050,-33.100,76.800,0.0000,0.0000,-150.0000
C00566=-23.050,-28.100,76.800,0.0000,0.0000,-150.0000
C00567=-23.050,-23.100,76.800,0.0000,0.0000,-150.0000
C00568=-23.050,-18.100,76.800,0.0000,0.0000,-150.0000
C00569=-23.050,-13.100,76.800,0.0000,0.0000,-150.0000
C00570=-23.050,-8.100,76.800,0.0000,0.0000,-150.0000
C00571=-23.050,-3.100,76.800,0.0000,0.0000,-150.0000
C00572=-23.050,1.900,76.800,0.0000,0.0000,-150.0000
C00573=-23.050,6.900,76.800,0.0000,0.0000,-150.0000
C00574=-23.050,11.900,76.800,0.0000,0.0000,-150.0000
C00575=-23.050,16.900,76.800,0.0000,0.0000,-150.0000
C00576=-23.050,21.900,76.800,0.0000,0.0000,-150.0000
C00577=-23.050,26.900,76.800,0.0000,0.0000,-150.0000
C00578=-23.050,31.900,76.800,0.0000,0.0000,-150.0000
C00579=-23.050,36.900,76.800,0.0000,0.0000,-150.0000
C00580=-23.050,41.900,76.800,0.0000,0.0000,-150.0000
C00581=-18.267,41.900,76.800,0.0000,0.0000,-150.0000
C00582=-13.483,41.900,76.800,0.0000,0.0000,-150.0000
C00583=-8.700,41.900,76.800,0.0000,0.0000,-150.0000
C00584=-3.917,41.900,76.800,0.0000,0.0000,-150.0000
C00585=0.867,41.900,76.800,0.0000,0.0000,-150.0000
C00586=5.650,41.900,76.800,0.0000,0.0000,-150.0000
C00587=10.433,41.900,76.800,0.0000,0.0000,-150.0000
C00588=15.217,41.900,76.800,0.0000,0.0000,-150.0000
C00589=20.000,41.900,76.800,0.0000,0.0000,-150.0000
C00590=25.000,41.900,76.800,0.0000,0.0000,-150.0000
C00591=26.950,43.850,76.800,0.0000,0.0000,-150.0000
C00592=25.000,45.800,76.800,0.0000,0.0000,-150.0000
C00593=20.000,45.800,76.800,0.0000,0.0000,-150.0000
C00594=15.000,45.800,76.800,0.0000,0.0000,-150.0000
C00595=10.000,45.800,76.800,0.0000,0.0000,-150.0000
C00596=5.000,45.800,76.800,0.0000,0.0000,-150.0000
C00597=0.000,45.800,76.800,0.0000,0.0000,-150.0000
C00598=-5.000,45.800,76.800,0.0000,0.0000,-150.0000
C00599=-10.000,45.800,76.800,0.0000,0.0000,-150.0000
C00600=-15.000,45.800,76.800,0.0000,0.0000,-150.0000
C00601=-20.000,45.800,76.800,0.0000,0.0000,-150.0000
C00602=-25.000,45.800,76.800,0.0000,0.0000,-150.0000
C00603=-30.000,45.800,76.800,0.0000,0.0000,-150.0000
C00604=-35.000,45.800,76.800,0.0000,0.0000,-150.0000
C00605=-40.000,45.800,76.800,0.0000,0.0000,-150.0000
C00606=-45.000,45.800,76.800,0.0000,0.0000,-150.0000
C00607=-50.000,45.800,76.800,0.0000,0.0000,-150.0000
C00608=-55.000,45.800,76.800,0.0000,0.0000,-150.0000
C00609=-60.000,45.800,76.800,0.0000,0.0000,-150.0000
C00610=-65.000,45.800,76.800,0.0000,0.0000,-150.0000
C00611=-70.000,45.800,76.800,0.0000,0.0000,-150.0000
C00612=-75.000,45.800,76.800,0.0000,0.0000,-150.0000
C00613=-76.950,43.850,76.800,0.0000,0.0000,-150.0000
C00614=-75.000,41.900,76.800,0.0000,0.0000,-150.0000
C00615=-70.195,41.900,76.800,0.0000,0.0000,-150.0000
C00616=-65.390,41.900,76.800,0.0000,0.0000,-150.0000
C00617=-60.585,41.900,76.800,0.0000,0.0000,-150.0000
C00618=-55.780,41.900,76.800,0.0000,0.0000,-150.0000
C00619=-50.975,41.900,76.800,0.0000,0.0000,-150.0000
C00620=-46.170,41.900,76.800,0.0000,0.0000,-150.0000
C00621=-41.365,41.900,76.800,0.0000,0.0000,-150.0000
C00622=-36.560,41.900,76.800,0.0000,0.0000,-150.0000
C00623=-31.755,41.900,76.800,0.0000,0.0000,-150.0000
C00624=-26.950,41.900,76.800,0.0000,0.0000,-150.0000
C00625=-26.950,36.900,76.800,0.0000,0.0000,-150.0000
C00626=-26.950,31.900,76.800,0.0000,0.0000,-150.0000
C00627=-26.950,26.900,76.800,0.0000,0.0000,-150.0000
C00628=-26.950,21.900,76.800,0.0000,0.0000,-150.0000
C00629=-26.950,16.900,76.800,0.0000,0.0000,-150.0000
C00630=-26.950,11.900,76.800,0.0000,0.0000,-150.0000
C00631=-26.950,6.900,76.800,0.0000,0.0000,-150.0000
C00632=-26.950,1.900,76.800,0.0000,0.0000,-150.0000
C00633=-26.950,-3.100,76.800,0.0000,0.0000,-150.0000
C00634=-26.950,-8.100,76.800,0.0000,0.0000,-150.0000
C00635=-26.950,-13.100,76.800,0.0000,0.0000,-150.0000
C00636=-26.950,-18.100,76.800,0.0000,0.0000,-150.0000
C00637=-26.950,-23.100,76.800,0.0000,0.0000,-150.0000
C00638=-26.950,-28.100,76.800,0.0000,0.0000,-150.0000
C00639=-26.950,-33.100,76.800,0.0000,0.0000,-150.0000
C00640=-26.950,-38.100,76.800,0.0000,0.0000,-150.0000
C00641=-26.950,-43.100,76.800,0.0000,0.0000,-150.0000
C00642=-26.950,-48.100,76.800,0.0000,0.0000,-150.0000
C00643=-26.950,-53.100,76.800,0.0000,0.0000,-150.0000
C00644=-26.950,-58.100,76.800,0.0000,0.0000,-150.0000
C00645=-26.950,-63.100,76.800,0.0000,0.0000,-150.0000
C00646=-26.950,-68.100,76.800,0.0000,0.0000,-150.0000
C00647=-31.755,-68.100,76.800,0.0000,0.0000,-150.0000
C00648=-36.560,-68.100,76.800,0.0000,0.0000,-150.0000
C00649=-41.365,-68.100,76.800,0.0000,0.0000,-150.0000
C00650=-46.170,-68.100,76.800,0.0000,0.0000,-150.0000
C00651=-50.975,-68.100,76.800,0.0000,0.0000,-150.0000
C00652=-55.780,-68.100,76.800,0.0000,0.0000,-150.0000
C00653=-60.585,-68.100,76.800,0.0000,0.0000,-150.0000
C00654=-65.390,-68.100,76.800,0.0000,0.0000,-150.0000
C00655=-70.195,-68.100,76.800,0.0000,0.0000,-150.0000
C00656=-75.000,-68.100,76.800,0.0000,0.0000,-150.0000
C00657=-75.000,-68.100,78.500,0.0000,0.0000,-150.0000
C00658=-70.195,-68.100,78.500,0.0000,0.0000,-150.0000
C00659=-65.390,-68.100,78.500,0.0000,0.0000,-150.0000
C00660=-60.585,-68.100,78.500,0.0000,0.0000,-150.0000
C00661=-55.780,-68.100,78.500,0.0000,0.0000,-150.0000
C00662=-50.975,-68.100,78.500,0.0000,0.0000,-150.0000
C00663=-46.170,-68.100,78.500,0.0000,0.0000,-150.0000
C00664=-41.365,-68.100,78.500,0.0000,0.0000,-150.0000
C00665=-36.560,-68.100,78.500,0.0000,0.0000,-150.0000
C00666=-31.755,-68.100,78.500,0.0000,0.0000,-150.0000
C00667=-26.950,-68.100,78.500,0.0000,0.0000,-150.0000
C00668=-26.950,-63.100,78.500,0.0000,0.0000,-150.0000
C00669=-26.950,-58.100,78.500,0.0000,0.0000,-150.0000
C00670=-26.950,-53.100,78.500,0.0000,0.0000,-150.0000
C00671=-26.950,-48.100,78.500,0.0000,0.0000,-150.0000
C00672=-26.950,-43.100,78.500,0.0000,0.0000,-150.0000
C00673=-26.950,-38.100,78.500,0.0000,0.0000,-150.0000
C00674=-26.950,-33.100,78.500,0.0000,0.0000,-150.0000
C00675=-26.950,-28.100,78.500,0.0000,0.0000,-150.0000
C00676=-26.950,-23.100,78.500,0.0000,0.0000,-150.0000
C00677=-26.950,-18.100,78.500,0.0000,0.0000,-150.0000
C00678=-26.950,-13.100,78.500,0.0000,0.0000,-150.0000
C00679=-26.950,-8.100,78.500,0.0000,0.0000,-150.0000
C00680=-26.950,-3.100,78.500,0.0000,0.0000,-150.0000
C00681=-26.950,1.900,78.500,0.0000,0.0000,-150.0000
C00682=-26.950,6.900,78.500,0.0000,0.0000,-150.0000
C00683=-26.950,11.900,78.500,0.0000,0.0000,-150.0000
C00684=-26.950,16.900,78.500,0.0000,0.0000,-150.0000
C00685=-26.950,21.900,78.500,0.0000,0.0000,-150.0000
C00686=-26.950,26.900,78.500,0.0000,0.0000,-150.0000
C00687=-26.950,31.900,78.500,0.0000,0.0000,-150.0000
C00688=-26.950,36.900,78.500,0.0000,0.0000,-150.0000
C00689=-26.950,41.900,78.500,0.0000,0.0000,-150.0000
C00690=-31.733,41.900,78.500,0.0000,0.0000,-150.0000
C00691=-36.517,41.900,78.500,0.0000,0.0000,-150.0000
C00692=-41.300,41.900,78.500,0.0000,0.0000,-150.0000
C00693=-46.083,41.900,78.500,0.0000,0.0000,-150.0000
C00694=-50.867,41.900,78.500,0.0000,0.0000,-150.0000
C00695=-55.650,41.900,78.500,0.0000,0.0000,-150.0000
C00696=-60.433,41.900,78.500,0.0000,0.0000,-150.0000
C00697=-65.217,41.900,78.500,0.0000,0.0000,-150.0000
C00698=-70.000,41.900,78.500,0.0000,0.0000,-150.0000
C00699=-75.000,41.900,78.500,0.0000,0.0000,-150.0000
C00700=-76.950,43.850,78.500,0.0000,0.0000,-150.0000
C00701=-75.000,45.800,78.500,0.0000,0.0000,-150.0000
C00702=-70.000,45.800,78.500,0.0000,0.0000,-150.0000
C00703=-65.000,45.800,78.500,0.0000,0.0000,-150.0000
C00704=-60.000,45.800,78.500,0.0000,0.0000,-150.0000
C00705=-55.000,45.800,78.500,0.0000,0.0000,-150.0000
C00706=-50.000,45.800,78.500,0.0000,0.0000,-150.0000
C00707=-45.000,45.800,78.500,0.0000,0.0000,-150.0000
C00708=-40.000,45.800,78.500,0.0000,0.0000,-150.0000
C00709=-35.000,45.800,78.500,0.0000,0.0000,-150.0000
C00710=-30.000,45.800,78.500,0.0000,0.0000,-150.0000
C00711=-25.000,45.800,78.500,0.0000,0.0000,-150.0000
C00712=-20.000,45.800,78.500,0.0000,0.0000,-150.0000
C00713=-15.000,45.800,78.500,0.0000,0.0000,-150.0000
C00714=-10.000,45.800,78.500,0.0000,0.0000,-150.0000
C00715=-5.000,45.800,78.500,0.0000,0.0000,-150.0000
C00716=0.000,45.800,78.500,0.0000,0.0000,-150.0000
C00717=5.000,45.800,78.500,0.0000,0.0000,-150.0000
C00718=10.000,45.800,78.500,0.0000,0.0000,-150.0000
C00719=15.000,45.800,78.500,0.0000,0.0000,-150.0000
C00720=20.000,45.800,78.500,0.0000,0.0000,-150.0000
C00721=25.000,45.800,78.500,0.0000,0.0000,-150.0000
C00722=26.950,43.850,78.500,0.0000,0.0000,-150.0000
C00723=25.000,41.900,78.500,0.0000,0.0000,-150.0000
C00724=20.195,41.900,78.500,0.0000,0.0000,-150.0000
C00725=15.390,41.900,78.500,0.0000,0.0000,-150.0000
C00726=10.585,41.900,78.500,0.0000,0.0000,-150.0000
C00727=5.780,41.900,78.500,0.0000,0.0000,-150.0000
C00728=0.975,41.900,78.500,0.0000,0.0000,-150.0000
C00729=-3.830,41.900,78.500,0.0000,0.0000,-150.0000
C00730=-8.635,41.900,78.500,0.0000,0.0000,-150.0000
C00731=-13.440,41.900,78.500,0.0000,0.0000,-150.0000
C00732=-18.245,41.900,78.500,0.0000,0.0000,-150.0000
C00733=-23.050,41.900,78.500,0.0000,0.0000,-150.0000
C00734=-23.050,36.900,78.500,0.0000,0.0000,-150.0000
C00735=-23.050,31.900,78.500,0.0000,0.0000,-150.0000
C00736=-23.050,26.900,78.500,0.0000,0.0000,-150.0000
C00737=-23.050,21.900,78.500,0.0000,0.0000,-150.0000
C00738=-23.050,16.900,78.500,0.0000,0.0000,-150.0000
C00739=-23.050,11.900,78.500,0.0000,0.0000,-150.0000
C00740=-23.050,6.900,78.500,0.0000,0.0000,-150.0000
C00741=-23.050,1.900,78.500,0.0000,0.0000,-150.0000
C00742=-23.050,-3.100,78.500,0.0000,0.0000,-150.0000
C00743=-23.050,-8.100,78.500,0.0000,0.0000,-150.0000
C00744=-23.050,-13.100,78.500,0.0000,0.0000,-150.0000
C00745=-23.050,-18.100,78.500,0.0000,0.0000,-150.0000
C00746=-23.050,-23.100,78.500,0.0000,0.0000,-150.0000
C00747=-23.050,-28.100,78.500,0.0000,0.0000,-150.0000
C00748=-23.050,-33.100,78.500,0.0000,0.0000,-150.0000
C00749=-23.050,-38.100,78.500,0.0000,0.0000,-150.0000
C00750=-23.050,-43.100,78.500,0.0000,0.0000,-150.0000
C00751=-23.050,-48.100,78.500,0.0000,0.0000,-150.0000
C00752=-23.050,-53.100,78.500,0.0000,0.0000,-150.0000
C00753=-23.050,-58.100,78.500,0.0000,0.0000,-150.0000
C00754=-23.050,-63.100,78.500,0.0000,0.0000,-150.0000
C00755=-23.050,-68.100,78.500,0.0000,0.0000,-150.0000
C00756=-18.267,-68.100,78.500,0.0000,0.0000,-150.0000
C00757=-13.483,-68.100,78.500,0.0000,0.0000,-150.0000
C00758=-8.700,-68.100,78.500,0.0000,0.0000,-150.0000
C00759=-3.917,-68.100,78.500,0.0000,0.0000,-150.0000
C00760=0.867,-68.100,78.500,0.0000,0.0000,-150.0000
C00761=5.650,-68.100,78.500,0.0000,0.0000,-150.0000
C00762=10.433,-68.100,78.500,0.0000,0.0000,-150.0000
C00763=15.217,-68.100,78.500,0.0000,0.0000,-150.0000
C00764=20.000,-68.100,78.500,0.0000,0.0000,-150.0000
C00765=25.000,-68.100,78.500,0.0000,0.0000,-150.0000
C00766=26.950,-70.050,78.500,0.0000,0.0000,-150.0000
C00767=25.000,-72.000,78.500,0.0000,0.0000,-150.0000
C00768=20.000,-72.000,78.500,0.0000,0.0000,-150.0000
C00769=15.000,-72.000,78.500,0.0000,0.0000,-150.0000
C00770=10.000,-72.000,78.500,0.0000,0.0000,-150.0000
C00771=5.000,-72.000,78.500,0.0000,0.0000,-150.0000
C00772=0.000,-72.000,78.500,0.0000,0.0000,-150.0000
C00773=-5.000,-72.000,78.500,0.0000,0.0000,-150.0000
C00774=-10.000,-72.000,78.500,0.0000,0.0000,-150.0000
C00775=-15.000,-72.000,78.500,0.0000,0.0000,-150.0000
C00776=-20.000,-72.000,78.500,0.0000,0.0000,-150.0000
C00777=-25.000,-72.000,78.500,0.0000,0.0000,-150.0000
C00778=-30.000,-72.000,78.500,0.0000,0.0000,-150.0000
C00779=-35.000,-72.000,78.500,0.0000,0.0000,-150.0000
C00780=-40.000,-72.000,78.500,0.0000,0.0000,-150.0000
C00781=-45.000,-72.000,78.500,0.0000,0.0000,-150.0000
C00782=-50.000,-72.000,78.500,0.0000,0.0000,-150.0000
C00783=-55.000,-72.000,78.500,0.0000,0.0000,-150.0000
C00784=-60.000,-72.000,78.500,0.0000,0.0000,-150.0000
C00785=-65.000,-72.000,78.500,0.0000,0.0000,-150.0000
C00786=-70.000,-72.000,78.500,0.0000,0.0000,-150.0000
C00787=-75.000,-72.000,78.500,0.0000,0.0000,-150.0000
C00788=-75.000,-72.000,80.200,0.0000,0.0000,-150.0000
C00789=-70.000,-72.000,80.200,0.0000,0.0000,-150.0000
C00790=-65.000,-72.000,80.200,0.0000,0.0000,-150.0000
C00791=-60.000,-72.000,80.200,0.0000,0.0000,-150.0000
C00792=-55.000,-72.000,80.200,0.0000,0.0000,-150.0000
C00793=-50.000,-72.000,80.200,0.0000,0.0000,-150.0000
C00794=-45.000,-72.000,80.200,0.0000,0.0000,-150.0000
C00795=-40.000,-72.000,80.200,0.0000,0.0000,-150.0000
C00796=-35.000,-72.000,80.200,0.0000,0.0000,-150.0000
C00797=-30.000,-72.000,80.200,0.0000,0.0000,-150.0000
C00798=-25.000,-72.000,80.200,0.0000,0.0000,-150.0000
C00799=-20.000,-72.000,80.200,0.0000,0.0000,-150.0000
C00800=-15.000,-72.000,80.200,0.0000,0.0000,-150.0000
C00801=-10.000,-72.000,80.200,0.0000,0.0000,-150.0000
C00802=-5.000,-72.000,80.200,0.0000,0.0000,-150.0000
C00803=0.000,-72.000,80.200,0.0000,0.0000,-150.0000
C00804=5.000,-72.000,80.200,0.0000,0.0000,-150.0000
C00805=10.000,-72.000,80.200,0.0000,0.0000,-150.0000
C00806=15.000,-72.000,80.200,0.0000,0.0000,-150.0000
C00807=20.000,-72.000,80.200,0.0000,0.0000,-150.0000
C00808=25.000,-72.000,80.200,0.0000,0.0000,-150.0000
C00809=26.950,-70.050,80.200,0.0000,0.0000,-150.0000
C00810=25.000,-68.100,80.200,0.0000,0.0000,-150.0000
C00811=20.195,-68.100,80.200,0.0000,0.0000,-150.0000
C00812=15.390,-68.100,80.200,0.0000,0.0000,-150.0000
C00813=10.585,-68.100,80.200,0.0000,0.0000,-150.0000
C00814=5.780,-68.100,80.200,0.0000,0.0000,-150.0000
C00815=0.975,-68.100,80.200,0.0000,0.0000,-150.0000
C00816=-3.830,-68.100,80.200,0.0000,0.0000,-150.0000
C00817=-8.635,-68.100,80.200,0.0000,0.0000,-150.0000
C00818=-13.440,-68.100,80.200,0.0000,0.0000,-150.0000
C00819=-18.245,-68.100,80.200,0.0000,0.0000,-150.0000
C00820=-23.050,-68.100,80.200,0.0000,0.0000,-150.0000
C00821=-23.050,-63.100,80.200,0.0000,0.0000,-150.0000
C00822=-23.050,-58.100,80.200,0.0000,0.0000,-150.0000
C00823=-23.050,-53.100,80.200,0.0000,0.0000,-150.0000
C00824=-23.050,-48.100,80.200,0.0000,0.0000,-150.0000
C00825=-23.050,-43.100,80.200,0.0000,0.0000,-150.0000
C00826=-23.050,-38.100,80.200,0.0000,0.0000,-150.0000
C00827=-23.050,-33.100,80.200,0.0000,0.0000,-150.0000
C00828=-23.050,-28.100,80.200,0.0000,0.0000,-150.0000
C00829=-23.050,-23.100,80.200,0.0000,0.0000,-150.0000
C00830=-23.050,-18.100,80.200,0.0000,0.0000,-150.0000
C00831=-23.050,-13.100,80.200,0.0000,0.0000,-150.0000
C00832=-23.050,-8.100,80.200,0.0000,0.0000,-150.0000
C00833=-23.050,-3.100,80.200,0.0000,0.0000,-150.0000
C00834=-23.050,1.900,80.200,0.0000,0.0000,-150.0000
C00835=-23.050,6.900,80.200,0.0000,0.0000,-150.0000
C00836=-23.050,11.900,80.200,0.0000,0.0000,-150.0000
C00837=-23.050,16.900,80.200,0.0000,0.0000,-150.0000
C00838=-23.050,21.900,80.200,0.0000,0.0000,-150.0000
C00839=-23.050,26.900,80.200,0.0000,0.0000,-150.0000
C00840=-23.050,31.900,80.200,0.0000,0.0000,-150.0000
C00841=-23.050,36.900,80.200,0.0000,0.0000,-150.0000
C00842=-23.050,41.900,80.200,0.0000,0.0000,-150.0000
C00843=-18.267,41.900,80.200,0.0000,0.0000,-150.0000
C00844=-13.483,41.900,80.200,0.0000,0.0000,-150.0000
C00845=-8.700,41.900,80.200,0.0000,0.0000,-150.0000
C00846=-3.917,41.900,80.200,0.0000,0.0000,-150.0000
C00847=0.867,41.900,80.200,0.0000,0.0000,-150.0000
C00848=5.650,41.900,80.200,0.0000,0.0000,-150.0000
C00849=10.433,41.900,80.200,0.0000,0.0000,-150.0000
C00850=15.217,41.900,80.200,0.0000,0.0000,-150.0000
C00851=20.000,41.900,80.200,0.0000,0.0000,-150.0000
C00852=25.000,41.900,80.200,0.0000,0.0000,-150.0000
C00853=26.950,43.850,80.200,0.0000,0.0000,-150.0000
C00854=25.000,45.800,80.200,0.0000,0.0000,-150.0000
C00855=20.000,45.800,80.200,0.0000,0.0000,-150.0000
C00856=15.000,45.800,80.200,0.0000,0.0000,-150.0000
C00857=10.000,45.800,80.200,0.0000,0.0000,-150.0000
C00858=5.000,45.800,80.200,0.0000,0.0000,-150.0000
C00859=0.000,45.800,80.200,0.0000,0.0000,-150.0000
C00860=-5.000,45.800,80.200,0.0000,0.0000,-150.0000
C00861=-10.000,45.800,80.200,0.0000,0.0000,-150.0000
C00862=-15.000,45.800,80.200,0.0000,0.0000,-150.0000
C00863=-20.000,45.800,80.200,0.0000,0.0000,-150.0000
C00864=-25.000,45.800,80.200,0.0000,0.0000,-150.0000
C00865=-30.000,45.800,80.200,0.0000,0.0000,-150.0000
C00866=-35.000,45.800,80.200,0.0000,0.0000,-150.0000
C00867=-40.000,45.800,80.200,0.0000,0.0000,-150.0000
C00868=-45.000,45.800,80.200,0.0000,0.0000,-150.0000
C00869=-50.000,45.800,80.200,0.0000,0.0000,-150.0000
C00870=-55.000,45.800,80.200,0.0000,0.0000,-150.0000
C00871=-60.000,45.800,80.200,0.0000,0.0000,-150.0000
C00872=-65.000,45.800,80.200,0.0000,0.0000,-150.0000
C00873=-70.000,45.800,80.200,0.0000,0.0000,-150.0000
C00874=-75.000,45.800,80.200,0.0000,0.0000,-150.0000
C00875=-76.950,43.850,80.200,0.0000,0.0000,-150.0000
C00876=-75.000,41.900,80.200,0.0000,0.0000,-150.0000
C00877=-70.195,41.900,80.200,0.0000,0.0000,-150.0000
C00878=-65.390,41.900,80.200,0.0000,0.0000,-150.0000
C00879=-60.585,41.900,80.200,0.0000,0.0000,-150.0000
C00880=-55.780,41.900,80.200,0.0000,0.0000,-150.0000
C00881=-50.975,41.900,80.200,0.0000,0.0000,-150.0000
C00882=-46.170,41.900,80.200,0.0000,0.0000,-150.0000
C00883=-41.365,41.900,80.200,0.0000,0.0000,-150.0000
C00884=-36.560,41.900,80.200,0.0000,0.0000,-150.0000
C00885=-31.755,41.900,80.200,0.0000,0.0000,-150.0000
C00886=-26.950,41.900,80.200,0.0000,0.0000,-150.0000
C00887=-26.950,36.900,80.200,0.0000,0.0000,-150.0000
C00888=-26.950,31.900,80.200,0.0000,0.0000,-150.0000
C00889=-26.950,26.900,80.200,0.0000,0.0000,-150.0000
C00890=-26.950,21.900,80.200,0.0000,0.0000,-150.0000
C00891=-26.950,16.900,80.200,0.0000,0.0000,-150.0000
C00892=-26.950,11.900,80.200,0.0000,0.0000,-150.0000
C00893=-26.950,6.900,80.200,0.0000,0.0000,-150.0000
C00894=-26.950,1.900,80.200,0.0000,0.0000,-150.0000
C00895=-26.950,-3.100,80.200,0.0000,0.0000,-150.0000
C00896=-26.950,-8.100,80.200,0.0000,0.0000,-150.0000
C00897=-26.950,-13.100,80.200,0.0000,0.0000,-150.0000
C00898=-26.950,-18.100,80.200,0.0000,0.0000,-150.0000
C00899=-26.950,-23.100,80.200,0.0000,0.0000,-150.0000
C00900=-26.950,-28.100,80.200,0.0000,0.0000,-150.0000
C00901=-26.950,-33.100,80.200,0.0000,0.0000,-150.0000
C00902=-26.950,-38.100,80.200,0.0000,0.0000,-150.0000
C00903=-26.950,-43.100,80.200,0.0000,0.0000,-150.0000
C00904=-26.950,-48.100,80.200,0.0000,0.0000,-150.0000
C00905=-26.950,-53.100,80.200,0.0000,0.0000,-150.0000
C00906=-26.950,-58.100,80.200,0.0000,0.0000,-150.0000
C00907=-26.950,-63.100,80.200,0.0000,0.0000,-150.0000
C00908=-26.950,-68.100,80.200,0.0000,0.0000,-150.0000
C00909=-31.755,-68.100,80.200,0.0000,0.0000,-150.0000
C00910=-36.560,-68.100,80.200,0.0000,0.0000,-150.0000
C00911=-41.365,-68.100,80.200,0.0000,0.0000,-150.0000
C00912=-46.170,-68.100,80.200,0.0000,0.0000,-150.0000
C00913=-50.975,-68.100,80.200,0.0000,0.0000,-150.0000
C00914=-55.780,-68.100,80.200,0.0000,0.0000,-150.0000
C00915=-60.585,-68.100,80.200,0.0000,0.0000,-150.0000
C00916=-65.390,-68.100,80.200,0.0000,0.0000,-150.0000
C00917=-70.195,-68.100,80.200,0.0000,0.0000,-150.0000
C00918=-75.000,-68.100,80.200,0.0000,0.0000,-150.0000
C00919=-75.000,-68.100,81.900,0.0000,0.0000,-150.0000
C00920=-70.195,-68.100,81.900,0.0000,0.0000,-150.0000
C00921=-65.390,-68.100,81.900,0.0000,0.0000,-150.0000
C00922=-60.585,-68.100,81.900,0.0000,0.0000,-150.0000
C00923=-55.780,-68.100,81.900,0.0000,0.0000,-150.0000
C00924=-50.975,-68.100,81.900,0.0000,0.0000,-150.0000
C00925=-46.170,-68.100,81.900,0.0000,0.0000,-150.0000
C00926=-41.365,-68.100,81.900,0.0000,0.0000,-150.0000
C00927=-36.560,-68.100,81.900,0.0000,0.0000,-150.0000
C00928=-31.755,-68.100,81.900,0.0000,0.0000,-150.0000
C00929=-26.950,-68.100,81.900,0.0000,0.0000,-150.0000
C00930=-26.950,-63.100,81.900,0.0000,0.0000,-150.0000
C00931=-26.950,-58.100,81.900,0.0000,0.0000,-150.0000
C00932=-26.950,-53.100,81.900,0.0000,0.0000,-150.0000
C00933=-26.950,-48.100,81.900,0.0000,0.0000,-150.0000
C00934=-26.950,-43.100,81.900,0.0000,0.0000,-150.0000
C00935=-26.950,-38.100,81.900,0.0000,0.0000,-150.0000
C00936=-26.950,-33.100,81.900,0.0000,0.0000,-150.0000
C00937=-26.950,-28.100,81.900,0.0000,0.0000,-150.0000
C00938=-26.950,-23.100,81.900,0.0000,0.0000,-150.0000
C00939=-26.950,-18.100,81.900,0.0000,0.0000,-150.0000
C00940=-26.950,-13.100,81.900,0.0000,0.0000,-150.0000
C00941=-26.950,-8.100,81.900,0.0000,0.0000,-150.0000
C00942=-26.950,-3.100,81.900,0.0000,0.0000,-150.0000
C00943=-26.950,1.900,81.900,0.0000,0.0000,-150.0000
C00944=-26.950,6.900,81.900,0.0000,0.0000,-150.0000
C00945=-26.950,11.900,81.900,0.0000,0.0000,-150.0000
C00946=-26.950,16.900,81.900,0.0000,0.0000,-150.0000
C00947=-26.950,21.900,81.900,0.0000,0.0000,-150.0000
C00948=-26.950,26.900,81.900,0.0000,0.0000,-150.0000
C00949=-26.950,31.900,81.900,0.0000,0.0000,-150.0000
C00950=-26.950,36.900,81.900,0.0000,0.0000,-150.0000
C00951=-26.950,41.900,81.900,0.0000,0.0000,-150.0000
C00952=-31.733,41.900,81.900,0.0000,0.0000,-150.0000
C00953=-36.517,41.900,81.900,0.0000,0.0000,-150.0000
C00954=-41.300,41.900,81.900,0.0000,0.0000,-150.0000
C00955=-46.083,41.900,81.900,0.0000,0.0000,-150.0000
C00956=-50.867,41.900,81.900,0.0000,0.0000,-150.0000
C00957=-55.650,41.900,81.900,0.0000,0.0000,-150.0000
C00958=-60.433,41.900,81.900,0.0000,0.0000,-150.0000
C00959=-65.217,41.900,81.900,0.0000,0.0000,-150.0000
C00960=-70.000,41.900,81.900,0.0000,0.0000,-150.0000
C00961=-75.000,41.900,81.900,0.0000,0.0000,-150.0000
C00962=-76.950,43.850,81.900,0.0000,0.0000,-150.0000
C00963=-75.000,45.800,81.900,0.0000,0.0000,-150.0000
C00964=-70.000,45.800,81.900,0.0000,0.0000,-150.0000
C00965=-65.000,45.800,81.900,0.0000,0.0000,-150.0000
C00966=-60.000,45.800,81.900,0.0000,0.0000,-150.0000
C00967=-55.000,45.800,81.900,0.0000,0.0000,-150.0000
C00968=-50.000,45.800,81.900,0.0000,0.0000,-150.0000
C00969=-45.000,45.800,81.900,0.0000,0.0000,-150.0000
C00970=-40.000,45.800,81.900,0.0000,0.0000,-150.0000
C00971=-35.000,45.800,81.900,0.0000,0.0000,-150.0000
C00972=-30.000,45.800,81.900,0.0000,0.0000,-150.0000
C00973=-25.000,45.800,81.900,0.0000,0.0000,-150.0000
C00974=-20.000,45.800,81.900,0.0000,0.0000,-150.0000
C00975=-15.000,45.800,81.900,0.0000,0.0000,-150.0000
C00976=-10.000,45.800,81.900,0.0000,0.0000,-150.0000
C00977=-5.000,45.800,81.900,0.0000,0.0000,-150.0000
C00978=0.000,45.800,81.900,0.0000,0.0000,-150.0000
C00979=5.000,45.800,81.900,0.0000,0.0000,-150.0000
C00980=10.000,45.800,81.900,0.0000,0.0000,-150.0000
C00981=15.000,45.800,81.900,0.0000,0.0000,-150.0000
C00982=20.000,45.800,81.900,0.0000,0.0000,-150.0000
C00983=25.000,45.800,81.900,0.0000,0.0000,-150.0000
C00984=26.950,43.850,81.900,0.0000,0.0000,-150.0000
C00985=25.000,41.900,81.900,0.0000,0.0000,-150.0000
C00986=20.195,41.900,81.900,0.0000,0.0000,-150.0000
C00987=15.390,41.900,81.900,0.0000,0.0000,-150.0000
C00988=10.585,41.900,81.900,0.0000,0.0000,-150.0000
C00989=5.780,41.900,81.900,0.0000,0.0000,-150.0000
C00990=0.975,41.900,81.900,0.0000,0.0000,-150.0000
C00991=-3.830,41.900,81.900,0.0000,0.0000,-150.0000
C00992=-8.635,41.900,81.900,0.0000,0.0000,-150.0000
C00993=-13.440,41.900,81.900,0.0000,0.0000,-150.0000
C00994=-18.245,41.900,81.900,0.0000,0.0000,-150.0000
C00995=-23.050,41.900,81.900,0.0000,0.0000,-150.0000
C00996=-23.050,36.900,81.900,0.0000,0.0000,-150.0000
C00997=-23.050,31.900,81.900,0.0000,0.0000,-150.0000
C00998=-23.050,26.900,81.900,0.0000,0.0000,-150.0000
C00999=-23.050,21.900,81.900,0.0000,0.0000,-150.0000
C01000=-23.050,16.900,81.900,0.0000,0.0000,-150.0000
C01001=-23.050,11.900,81.900,0.0000,0.0000,-150.0000
C01002=-23.050,6.900,81.900,0.0000,0.0000,-150.0000
C01003=-23.050,1.900,81.900,0.0000,0.0000,-150.0000
C01004=-23.050,-3.100,81.900,0.0000,0.0000,-150.0000
C01005=-23.050,-8.100,81.900,0.0000,0.0000,-150.0000
C01006=-23.050,-13.100,81.900,0.0000,0.0000,-150.0000
C01007=-23.050,-18.100,81.900,0.0000,0.0000,-150.0000
C01008=-23.050,-23.100,81.900,0.0000,0.0000,-150.0000
C01009=-23.050,-28.100,81.900,0.0000,0.0000,-150.0000
C01010=-23.050,-33.100,81.900,0.0000,0.0000,-150.0000
C01011=-23.050,-38.100,81.900,0.0000,0.0000,-150.0000
C01012=-23.050,-43.100,81.900,0.0000,0.0000,-150.0000
C01013=-23.050,-48.100,81.900,0.0000,0.0000,-150.0000
C01014=-23.050,-53.100,81.900,0.0000,0.0000,-150.0000
C01015=-23.050,-58.100,81.900,0.0000,0.0000,-150.0000
C01016=-23.050,-63.100,81.900,0.0000,0.0000,-150.0000
C01017=-23.050,-68.100,81.900,0.0000,0.0000,-150.0000
C01018=-18.267,-68.100,81.900,0.0000,0.0000,-150.0000
C01019=-13.483,-68.100,81.900,0.0000,0.0000,-150.0000
C01020=-8.700,-68.100,81.900,0.0000,0.0000,-150.0000
C01021=-3.917,-68.100,81.900,0.0000,0.0000,-150.0000
C01022=0.867,-68.100,81.900,0.0000,0.0000,-150.0000
C01023=5.650,-68.100,81.900,0.0000,0.0000,-150.0000
C01024=10.433,-68.100,81.900,0.0000,0.0000,-150.0000
C01025=15.217,-68.100,81.900,0.0000,0.0000,-150.0000
C01026=20.000,-68.100,81.900,0.0000,0.0000,-150.0000
C01027=25.000,-68.100,81.900,0.0000,0.0000,-150.0000
C01028=26.950,-70.050,81.900,0.0000,0.0000,-150.0000
C01029=25.000,-72.000,81.900,0.0000,0.0000,-150.0000
C01030=20.000,-72.000,81.900,0.0000,0.0000,-150.0000
C01031=15.000,-72.000,81.900,0.0000,0.0000,-150.0000
C01032=10.000,-72.000,81.900,0.0000,0.0000,-150.0000
C01033=5.000,-72.000,81.900,0.0000,0.0000,-150.0000
C01034=0.000,-72.000,81.900,0.0000,0.0000,-150.0000
C01035=-5.000,-72.000,81.900,0.0000,0.0000,-150.0000
C01036=-10.000,-72.000,81.900,0.0000,0.0000,-150.0000
C01037=-15.000,-72.000,81.900,0.0000,0.0000,-150.0000
C01038=-20.000,-72.000,81.900,0.0000,0.0000,-150.0000
C01039=-25.000,-72.000,81.900,0.0000,0.0000,-150.0000
C01040=-30.000,-72.000,81.900,0.0000,0.0000,-150.0000
C01041=-35.000,-72.000,81.900,0.0000,0.0000,-150.0000
C01042=-40.000,-72.000,81.900,0.0000,0.0000,-150.0000
C01043=-45.000,-72.000,81.900,0.0000,0.0000,-150.0000
C01044=-50.000,-72.000,81.900,0.0000,0.0000,-150.0000
C01045=-55.000,-72.000,81.900,0.0000,0.0000,-150.0000
C01046=-60.000,-72.000,81.900,0.0000,0.0000,-150.0000
C01047=-65.000,-72.000,81.900,0.0000,0.0000,-150.0000
C01048=-70.000,-72.000,81.900,0.0000,0.0000,-150.0000
C01049=-75.000,-72.000,81.900,0.0000,0.0000,-150.0000
C01050=-75.000,-72.000,83.600,0.0000,0.0000,-150.0000
C01051=-70.000,-72.000,83.600,0.0000,0.0000,-150.0000
C01052=-65.000,-72.000,83.600,0.0000,0.0000,-150.0000
C01053=-60.000,-72.000,83.600,0.0000,0.0000,-150.0000
C01054=-55.000,-72.000,83.600,0.0000,0.0000,-150.0000
C01055=-50.000,-72.000,83.600,0.0000,0.0000,-150.0000
C01056=-45.000,-72.000,83.600,0.0000,0.0000,-150.0000
C01057=-40.000,-72.000,83.600,0.0000,0.0000,-150.0000
C01058=-35.000,-72.000,83.600,0.0000,0.0000,-150.0000
C01059=-30.000,-72.000,83.600,0.0000,0.0000,-150.0000
C01060=-25.000,-72.000,83.600,0.0000,0.0000,-150.0000
C01061=-20.000,-72.000,83.600,0.0000,0.0000,-150.0000
C01062=-15.000,-72.000,83.600,0.0000,0.0000,-150.0000
C01063=-10.000,-72.000,83.600,0.0000,0.0000,-150.0000
C01064=-5.000,-72.000,83.600,0.0000,0.0000,-150.0000
C01065=0.000,-72.000,83.600,0.0000,0.0000,-150.0000
C01066=5.000,-72.000,83.600,0.0000,0.0000,-150.0000
C01067=10.000,-72.000,83.600,0.0000,0.0000,-150.0000
C01068=15.000,-72.000,83.600,0.0000,0.0000,-150.0000
C01069=20.000,-72.000,83.600,0.0000,0.0000,-150.0000
C01070=25.000,-72.000,83.600,0.0000,0.0000,-150.0000
C01071=26.950,-70.050,83.600,0.0000,0.0000,-150.0000
C01072=25.000,-68.100,83.600,0.0000,0.0000,-150.0000
C01073=20.195,-68.100,83.600,0.0000,0.0000,-150.0000
C01074=15.390,-68.100,83.600,0.0000,0.0000,-150.0000
C01075=10.585,-68.100,83.600,0.0000,0.0000,-150.0000
C01076=5.780,-68.100,83.600,0.0000,0.0000,-150.0000
C01077=0.975,-68.100,83.600,0.0000,0.0000,-150.0000
C01078=-3.830,-68.100,83.600,0.0000,0.0000,-150.0000
C01079=-8.635,-68.100,83.600,0.0000,0.0000,-150.0000
C01080=-13.440,-68.100,83.600,0.0000,0.0000,-150.0000
C01081=-18.245,-68.100,83.600,0.0000,0.0000,-150.0000
C01082=-23.050,-68.100,83.600,0.0000,0.0000,-150.0000
C01083=-23.050,-63.100,83.600,0.0000,0.0000,-150.0000
C01084=-23.050,-58.100,83.600,0.0000,0.0000,-150.0000
C01085=-23.050,-53.100,83.600,0.0000,0.0000,-150.0000
C01086=-23.050,-48.100,83.600,0.0000,0.0000,-150.0000
C01087=-23.050,-43.100,83.600,0.0000,0.0000,-150.0000
C01088=-23.050,-38.100,83.600,0.0000,0.0000,-150.0000
C01089=-23.050,-33.100,83.600,0.0000,0.0000,-150.0000
C01090=-23.050,-28.100,83.600,0.0000,0.0000,-150.0000
C01091=-23.050,-23.100,83.600,0.0000,0.0000,-150.0000
C01092=-23.050,-18.100,83.600,0.0000,0.0000,-150.0000
C01093=-23.050,-13.100,83.600,0.0000,0.0000,-150.0000
C01094=-23.050,-8.100,83.600,0.0000,0.0000,-150.0000
C01095=-23.050,-3.100,83.600,0.0000,0.0000,-150.0000
C01096=-23.050,1.900,83.600,0.0000,0.0000,-150.0000
C01097=-23.050,6.900,83.600,0.0000,0.0000,-150.0000
C01098=-23.050,11.900,83.600,0.0000,0.0000,-150.0000
C01099=-23.050,16.900,83.600,0.0000,0.0000,-150.0000
C01100=-23.050,21.900,83.600,0.0000,0.0000,-150.0000
C01101=-23.050,26.900,83.600,0.0000,0.0000,-150.0000
C01102=-23.050,31.900,83.600,0.0000,0.0000,-150.0000
C01103=-23.050,36.900,83.600,0.0000,0.0000,-150.0000
C01104=-23.050,41.900,83.600,0.0000,0.0000,-150.0000
C01105=-18.267,41.900,83.600,0.0000,0.0000,-150.0000
C01106=-13.483,41.900,83.600,0.0000,0.0000,-150.0000
C01107=-8.700,41.900,83.600,0.0000,0.0000,-150.0000
C01108=-3.917,41.900,83.600,0.0000,0.0000,-150.0000
C01109=0.867,41.900,83.600,0.0000,0.0000,-150.0000
C01110=5.650,41.900,83.600,0.0000,0.0000,-150.0000
C01111=10.433,41.900,83.600,0.0000,0.0000,-150.0000
C01112=15.217,41.900,83.600,0.0000,0.0000,-150.0000
C01113=20.000,41.900,83.600,0.0000,0.0000,-150.0000
C01114=25.000,41.900,83.600,0.0000,0.0000,-150.0000
C01115=26.950,43.850,83.600,0.0000,0.0000,-150.0000
C01116=25.000,45.800,83.600,0.0000,0.0000,-150.0000
C01117=20.000,45.800,83.600,0.0000,0.0000,-150.0000
C01118=15.000,45.800,83.600,0.0000,0.0000,-150.0000
C01119=10.000,45.800,83.600,0.0000,0.0000,-150.0000
C01120=5.000,45.800,83.600,0.0000,0.0000,-150.0000
C01121=0.000,45.800,83.600,0.0000,0.0000,-150.0000
C01122=-5.000,45.800,83.600,0.0000,0.0000,-150.0000
C01123=-10.000,45.800,83.600,0.0000,0.0000,-150.0000
C01124=-15.000,45.800,83.600,0.0000,0.0000,-150.0000
C01125=-20.000,45.800,83.600,0.0000,0.0000,-150.0000
C01126=-25.000,45.800,83.600,0.0000,0.0000,-150.0000
C01127=-30.000,45.800,83.600,0.0000,0.0000,-150.0000
C01128=-35.000,45.800,83.600,0.0000,0.0000,-150.0000
C01129=-40.000,45.800,83.600,0.0000,0.0000,-150.0000
C01130=-45.000,45.800,83.600,0.0000,0.0000,-150.0000
C01131=-50.000,45.800,83.600,0.0000,0.0000,-150.0000
C01132=-55.000,45.800,83.600,0.0000,0.0000,-150.0000
C01133=-60.000,45.800,83.600,0.0000,0.0000,-150.0000
C01134=-65.000,45.800,83.600,0.0000,0.0000,-150.0000
C01135=-70.000,45.800,83.600,0.0000,0.0000,-150.0000
C01136=-75.000,45.800,83.600,0.0000,0.0000,-150.0000
C01137=-76.950,43.850,83.600,0.0000,0.0000,-150.0000
C01138=-75.000,41.900,83.600,0.0000,0.0000,-150.0000
C01139=-70.195,41.900,83.600,0.0000,0.0000,-150.0000
C01140=-65.390,41.900,83.600,0.0000,0.0000,-150.0000
C01141=-60.585,41.900,83.600,0.0000,0.0000,-150.0000
C01142=-55.780,41.900,83.600,0.0000,0.0000,-150.0000
C01143=-50.975,41.900,83.600,0.0000,0.0000,-150.0000
C01144=-46.170,41.900,83.600,0.0000,0.0000,-150.0000
C01145=-41.365,41.900,83.600,0.0000,0.0000,-150.0000
C01146=-36.560,41.900,83.600,0.0000,0.0000,-150.0000
C01147=-31.755,41.900,83.600,0.0000,0.0000,-150.0000
C01148=-26.950,41.900,83.600,0.0000,0.0000,-150.0000
C01149=-26.950,36.900,83.600,0.0000,0.0000,-150.0000
C01150=-26.950,31.900,83.600,0.0000,0.0000,-150.0000
C01151=-26.950,26.900,83.600,0.0000,0.0000,-150.0000
C01152=-26.950,21.900,83.600,0.0000,0.0000,-150.0000
C01153=-26.950,16.900,83.600,0.0000,0.0000,-150.0000
C01154=-26.950,11.900,83.600,0.0000,0.0000,-150.0000
C01155=-26.950,6.900,83.600,0.0000,0.0000,-150.0000
C01156=-26.950,1.900,83.600,0.0000,0.0000,-150.0000
C01157=-26.950,-3.100,83.600,0.0000,0.0000,-150.0000
C01158=-26.950,-8.100,83.600,0.0000,0.0000,-150.0000
C01159=-26.950,-13.100,83.600,0.0000,0.0000,-150.0000
C01160=-26.950,-18.100,83.600,0.0000,0.0000,-150.0000
C01161=-26.950,-23.100,83.600,0.0000,0.0000,-150.0000
C01162=-26.950,-28.100,83.600,0.0000,0.0000,-150.0000
C01163=-26.950,-33.100,83.600,0.0000,0.0000,-150.0000
C01164=-26.950,-38.100,83.600,0.0000,0.0000,-150.0000
C01165=-26.950,-43.100,83.600,0.0000,0.0000,-150.0000
C01166=-26.950,-48.100,83.600,0.0000,0.0000,-150.0000
C01167=-26.950,-53.100,83.600,0.0000,0.0000,-150.0000
C01168=-26.950,-58.100,83.600,0.0000,0.0000,-150.0000
C01169=-26.950,-63.100,83.600,0.0000,0.0000,-150.0000
C01170=-26.950,-68.100,83.600,0.0000,0.0000,-150.0000
C01171=-31.755,-68.100,83.600,0.0000,0.0000,-150.0000
C01172=-36.560,-68.100,83.600,0.0000,0.0000,-150.0000
C01173=-41.365,-68.100,83.600,0.0000,0.0000,-150.0000
C01174=-46.170,-68.100,83.600,0.0000,0.0000,-150.0000
C01175=-50.975,-68.100,83.600,0.0000,0.0000,-150.0000
C01176=-55.780,-68.100,83.600,0.0000,0.0000,-150.0000
C01177=-60.585,-68.100,83.600,0.0000,0.0000,-150.0000
C01178=-65.390,-68.100,83.600,0.0000,0.0000,-150.0000
C01179=-70.195,-68.100,83.600,0.0000,0.0000,-150.0000
C01180=-75.000,-68.100,83.600,0.0000,0.0000,-150.0000
C01181=-75.000,-68.100,85.300,0.0000,0.0000,-150.0000
C01182=-70.195,-68.100,85.300,0.0000,0.0000,-150.0000
C01183=-65.390,-68.100,85.300,0.0000,0.0000,-150.0000
C01184=-60.585,-68.100,85.300,0.0000,0.0000,-150.0000
C01185=-55.780,-68.100,85.300,0.0000,0.0000,-150.0000
C01186=-50.975,-68.100,85.300,0.0000,0.0000,-150.0000
C01187=-46.170,-68.100,85.300,0.0000,0.0000,-150.0000
C01188=-41.365,-68.100,85.300,0.0000,0.0000,-150.0000
C01189=-36.560,-68.100,85.300,0.0000,0.0000,-150.0000
C01190=-31.755,-68.100,85.300,0.0000,0.0000,-150.0000
C01191=-26.950,-68.100,85.300,0.0000,0.0000,-150.0000
C01192=-26.950,-63.100,85.300,0.0000,0.0000,-150.0000
C01193=-26.950,-58.100,85.300,0.0000,0.0000,-150.0000
C01194=-26.950,-53.100,85.300,0.0000,0.0000,-150.0000
C01195=-26.950,-48.100,85.300,0.0000,0.0000,-150.0000
C01196=-26.950,-43.100,85.300,0.0000,0.0000,-150.0000
C01197=-26.950,-38.100,85.300,0.0000,0.0000,-150.0000
C01198=-26.950,-33.100,85.300,0.0000,0.0000,-150.0000
C01199=-26.950,-28.100,85.300,0.0000,0.0000,-150.0000
C01200=-26.950,-23.100,85.300,0.0000,0.0000,-150.0000
C01201=-26.950,-18.100,85.300,0.0000,0.0000,-150.0000
C01202=-26.950,-13.100,85.300,0.0000,0.0000,-150.0000
C01203=-26.950,-8.100,85.300,0.0000,0.0000,-150.0000
C01204=-26.950,-3.100,85.300,0.0000,0.0000,-150.0000
C01205=-26.950,1.900,85.300,0.0000,0.0000,-150.0000
C01206=-26.950,6.900,85.300,0.0000,0.0000,-150.0000
C01207=-26.950,11.900,85.300,0.0000,0.0000,-150.0000
C01208=-26.950,16.900,85.300,0.0000,0.0000,-150.0000
C01209=-26.950,21.900,85.300,0.0000,0.0000,-150.0000
C01210=-26.950,26.900,85.300,0.0000,0.0000,-150.0000
C01211=-26.950,31.900,85.300,0.0000,0.0000,-150.0000
C01212=-26.950,36.900,85.300,0.0000,0.0000,-150.0000
C01213=-26.950,41.900,85.300,0.0000,0.0000,-150.0000
C01214=-31.733,41.900,85.300,0.0000,0.0000,-150.0000
C01215=-36.517,41.900,85.300,0.0000,0.0000,-150.0000
C01216=-41.300,41.900,85.300,0.0000,0.0000,-150.0000
C01217=-46.083,41.900,85.300,0.0000,0.0000,-150.0000
C01218=-50.867,41.900,85.300,0.0000,0.0000,-150.0000
C01219=-55.650,41.900,85.300,0.0000,0.0000,-150.0000
C01220=-60.433,41.900,85.300,0.0000,0.0000,-150.0000
C01221=-65.217,41.900,85.300,0.0000,0.0000,-150.0000
C01222=-70.000,41.900,85.300,0.0000,0.0000,-150.0000
C01223=-75.000,41.900,85.300,0.0000,0.0000,-150.0000
C01224=-76.950,43.850,85.300,0.0000,0.0000,-150.0000
C01225=-75.000,45.800,85.300,0.0000,0.0000,-150.0000
C01226=-70.000,45.800,85.300,0.0000,0.0000,-150.0000
C01227=-65.000,45.800,85.300,0.0000,0.0000,-150.0000
C01228=-60.000,45.800,85.300,0.0000,0.0000,-150.0000
C01229=-55.000,45.800,85.300,0.0000,0.0000,-150.0000
C01230=-50.000,45.800,85.300,0.0000,0.0000,-150.0000
C01231=-45.000,45.800,85.300,0.0000,0.0000,-150.0000
C01232=-40.000,45.800,85.300,0.0000,0.0000,-150.0000
C01233=-35.000,45.800,85.300,0.0000,0.0000,-150.0000
C01234=-30.000,45.800,85.300,0.0000,0.0000,-150.0000
C01235=-25.000,45.800,85.300,0.0000,0.0000,-150.0000
C01236=-20.000,45.800,85.300,0.0000,0.0000,-150.0000
C01237=-15.000,45.800,85.300,0.0000,0.0000,-150.0000
C01238=-10.000,45.800,85.300,0.0000,0.0000,-150.0000
C01239=-5.000,45.800,85.300,0.0000,0.0000,-150.0000
C01240=0.000,45.800,85.300,0.0000,0.0000,-150.0000
C01241=5.000,45.800,85.300,0.0000,0.0000,-150.0000
C01242=10.000,45.800,85.300,0.0000,0.0000,-150.0000
C01243=15.000,45.800,85.300,0.0000,0.0000,-150.0000
C01244=20.000,45.800,85.300,0.0000,0.0000,-150.0000
C01245=25.000,45.800,85.300,0.0000,0.0000,-150.0000
C01246=26.950,43.850,85.300,0.0000,0.0000,-150.0000
C01247=25.000,41.900,85.300,0.0000,0.0000,-150.0000
C01248=20.195,41.900,85.300,0.0000,0.0000,-150.0000
C01249=15.390,41.900,85.300,0.0000,0.0000,-150.0000
C01250=10.585,41.900,85.300,0.0000,0.0000,-150.0000
C01251=5.780,41.900,85.300,0.0000,0.0000,-150.0000
C01252=0.975,41.900,85.300,0.0000,0.0000,-150.0000
C01253=-3.830,41.900,85.300,0.0000,0.0000,-150.0000
C01254=-8.635,41.900,85.300,0.0000,0.0000,-150.0000
C01255=-13.440,41.900,85.300,0.0000,0.0000,-150.0000
C01256=-18.245,41.900,85.300,0.0000,0.0000,-150.0000
C01257=-23.050,41.900,85.300,0.0000,0.0000,-150.0000
C01258=-23.050,36.900,85.300,0.0000,0.0000,-150.0000
C01259=-23.050,31.900,85.300,0.0000,0.0000,-150.0000
C01260=-23.050,26.900,85.300,0.0000,0.0000,-150.0000
C01261=-23.050,21.900,85.300,0.0000,0.0000,-150.0000
C01262=-23.050,16.900,85.300,0.0000,0.0000,-150.0000
C01263=-23.050,11.900,85.300,0.0000,0.0000,-150.0000
C01264=-23.050,6.900,85.300,0.0000,0.0000,-150.0000
C01265=-23.050,1.900,85.300,0.0000,0.0000,-150.0000
C01266=-23.050,-3.100,85.300,0.0000,0.0000,-150.0000
C01267=-23.050,-8.100,85.300,0.0000,0.0000,-150.0000
C01268=-23.050,-13.100,85.300,0.0000,0.0000,-150.0000
C01269=-23.050,-18.100,85.300,0.0000,0.0000,-150.0000
C01270=-23.050,-23.100,85.300,0.0000,0.0000,-150.0000
C01271=-23.050,-28.100,85.300,0.0000,0.0000,-150.0000
C01272=-23.050,-33.100,85.300,0.0000,0.0000,-150.0000
C01273=-23.050,-38.100,85.300,0.0000,0.0000,-150.0000
C01274=-23.050,-43.100,85.300,0.0000,0.0000,-150.0000
C01275=-23.050,-48.100,85.300,0.0000,0.0000,-150.0000
C01276=-23.050,-53.100,85.300,0.0000,0.0000,-150.0000
C01277=-23.050,-58.100,85.300,0.0000,0.0000,-150.0000
C01278=-23.050,-63.100,85.300,0.0000,0.0000,-150.0000
C01279=-23.050,-68.100,85.300,0.0000,0.0000,-150.0000
C01280=-18.267,-68.100,85.300,0.0000,0.0000,-150.0000
C01281=-13.483,-68.100,85.300,0.0000,0.0000,-150.0000
C01282=-8.700,-68.100,85.300,0.0000,0.0000,-150.0000
C01283=-3.917,-68.100,85.300,0.0000,0.0000,-150.0000
C01284=0.867,-68.100,85.300,0.0000,0.0000,-150.0000
C01285=5.650,-68.100,85.300,0.0000,0.0000,-150.0000
C01286=10.433,-68.100,85.300,0.0000,0.0000,-150.0000
C01287=15.217,-68.100,85.300,0.0000,0.0000,-150.0000
C01288=20.000,-68.100,85.300,0.0000,0.0000,-150.0000
C01289=25.000,-68.100,85.300,0.0000,0.0000,-150.0000
C01290=26.950,-70.050,85.300,0.0000,0.0000,-150.0000
C01291=25.000,-72.000,85.300,0.0000,0.0000,-150.0000
C01292=20.000,-72.000,85.300,0.0000,0.0000,-150.0000
C01293=15.000,-72.000,85.300,0.0000,0.0000,-150.0000
C01294=10.000,-72.000,85.300,0.0000,0.0000,-150.0000
C01295=5.000,-72.000,85.300,0.0000,0.0000,-150.0000
C01296=0.000,-72.000,85.300,0.0000,0.0000,-150.0000
C01297=-5.000,-72.000,85.300,0.0000,0.0000,-150.0000
C01298=-10.000,-72.000,85.300,0.0000,0.0000,-150.0000
C01299=-15.000,-72.000,85.300,0.0000,0.0000,-150.0000
C01300=-20.000,-72.000,85.300,0.0000,0.0000,-150.0000
C01301=-25.000,-72.000,85.300,0.0000,0.0000,-150.0000
C01302=-30.000,-72.000,85.300,0.0000,0.0000,-150.0000
C01303=-35.000,-72.000,85.300,0.0000,0.0000,-150.0000
C01304=-40.000,-72.000,85.300,0.0000,0.0000,-150.0000
C01305=-45.000,-72.000,85.300,0.0000,0.0000,-150.0000
C01306=-50.000,-72.000,85.300,0.0000,0.0000,-150.0000
C01307=-55.000,-72.000,85.300,0.0000,0.0000,-150.0000
C01308=-60.000,-72.000,85.300,0.0000,0.0000,-150.0000
C01309=-65.000,-72.000,85.300,0.0000,0.0000,-150.0000
C01310=-70.000,-72.000,85.300,0.0000,0.0000,-150.0000
C01311=-75.000,-72.000,85.300,0.0000,0.0000,-150.0000
C01312=-75.000,-72.000,87.000,0.0000,0.0000,-150.0000
C01313=-70.000,-72.000,87.000,0.0000,0.0000,-150.0000
C01314=-65.000,-72.000,87.000,0.0000,0.0000,-150.0000
C01315=-60.000,-72.000,87.000,0.0000,0.0000,-150.0000
C01316=-55.000,-72.000,87.000,0.0000,0.0000,-150.0000
C01317=-50.000,-72.000,87.000,0.0000,0.0000,-150.0000
C01318=-45.000,-72.000,87.000,0.0000,0.0000,-150.0000
C01319=-40.000,-72.000,87.000,0.0000,0.0000,-150.0000
C01320=-35.000,-72.000,87.000,0.0000,0.0000,-150.0000
C01321=-30.000,-72.000,87.000,0.0000,0.0000,-150.0000
C01322=-25.000,-72.000,87.000,0.0000,0.0000,-150.0000
C01323=-20.000,-72.000,87.000,0.0000,0.0000,-150.0000
C01324=-15.000,-72.000,87.000,0.0000,0.0000,-150.0000
C01325=-10.000,-72.000,87.000,0.0000,0.0000,-150.0000
C01326=-5.000,-72.000,87.000,0.0000,0.0000,-150.0000
C01327=0.000,-72.000,87.000,0.0000,0.0000,-150.0000
C01328=5.000,-72.000,87.000,0.0000,0.0000,-150.0000
C01329=10.000,-72.000,87.000,0.0000,0.0000,-150.0000
C01330=15.000,-72.000,87.000,0.0000,0.0000,-150.0000
C01331=20.000,-72.000,87.000,0.0000,0.0000,-150.0000
C01332=25.000,-72.000,87.000,0.0000,0.0000,-150.0000
C01333=26.950,-70.050,87.000,0.0000,0.0000,-150.0000
C01334=25.000,-68.100,87.000,0.0000,0.0000,-150.0000
C01335=20.195,-68.100,87.000,0.0000,0.0000,-150.0000
C01336=15.390,-68.100,87.000,0.0000,0.0000,-150.0000
C01337=10.585,-68.100,87.000,0.0000,0.0000,-150.0000
C01338=5.780,-68.100,87.000,0.0000,0.0000,-150.0000
C01339=0.975,-68.100,87.000,0.0000,0.0000,-150.0000
C01340=-3.830,-68.100,87.000,0.0000,0.0000,-150.0000
C01341=-8.635,-68.100,87.000,0.0000,0.0000,-150.0000
C01342=-13.440,-68.100,87.000,0.0000,0.0000,-150.0000
C01343=-18.245,-68.100,87.000,0.0000,0.0000,-150.0000
C01344=-23.050,-68.100,87.000,0.0000,0.0000,-150.0000
C01345=-23.050,-63.100,87.000,0.0000,0.0000,-150.0000
C01346=-23.050,-58.100,87.000,0.0000,0.0000,-150.0000
C01347=-23.050,-53.100,87.000,0.0000,0.0000,-150.0000
C01348=-23.050,-48.100,87.000,0.0000,0.0000,-150.0000
C01349=-23.050,-43.100,87.000,0.0000,0.0000,-150.0000
C01350=-23.050,-38.100,87.000,0.0000,0.0000,-150.0000
C01351=-23.050,-33.100,87.000,0.0000,0.0000,-150.0000
C01352=-23.050,-28.100,87.000,0.0000,0.0000,-150.0000
C01353=-23.050,-23.100,87.000,0.0000,0.0000,-150.0000
C01354=-23.050,-18.100,87.000,0.0000,0.0000,-150.0000
C01355=-23.050,-13.100,87.000,0.0000,0.0000,-150.0000
C01356=-23.050,-8.100,87.000,0.0000,0.0000,-150.0000
C01357=-23.050,-3.100,87.000,0.0000,0.0000,-150.0000
C01358=-23.050,1.900,87.000,0.0000,0.0000,-150.0000
C01359=-23.050,6.900,87.000,0.0000,0.0000,-150.0000
C01360=-23.050,11.900,87.000,0.0000,0.0000,-150.0000
C01361=-23.050,16.900,87.000,0.0000,0.0000,-150.0000
C01362=-23.050,21.900,87.000,0.0000,0.0000,-150.0000
C01363=-23.050,26.900,87.000,0.0000,0.0000,-150.0000
C01364=-23.050,31.900,87.000,0.0000,0.0000,-150.0000
C01365=-23.050,36.900,87.000,0.0000,0.0000,-150.0000
C01366=-23.050,41.900,87.000,0.0000,0.0000,-150.0000
C01367=-18.267,41.900,87.000,0.0000,0.0000,-150.0000
C01368=-13.483,41.900,87.000,0.0000,0.0000,-150.0000
C01369=-8.700,41.900,87.000,0.0000,0.0000,-150.0000
C01370=-3.917,41.900,87.000,0.0000,0.0000,-150.0000
C01371=0.867,41.900,87.000,0.0000,0.0000,-150.0000
C01372=5.650,41.900,87.000,0.0000,0.0000,-150.0000
C01373=10.433,41.900,87.000,0.0000,0.0000,-150.0000
C01374=15.217,41.900,87.000,0.0000,0.0000,-150.0000
C01375=20.000,41.900,87.000,0.0000,0.0000,-150.0000
C01376=25.000,41.900,87.000,0.0000,0.0000,-150.0000
C01377=26.950,43.850,87.000,0.0000,0.0000,-150.0000
C01378=25.000,45.800,87.000,0.0000,0.0000,-150.0000
C01379=20.000,45.800,87.000,0.0000,0.0000,-150.0000
C01380=15.000,45.800,87.000,0.0000,0.0000,-150.0000
C01381=10.000,45.800,87.000,0.0000,0.0000,-150.0000
C01382=5.000,45.800,87.000,0.0000,0.0000,-150.0000
C01383=0.000,45.800,87.000,0.0000,0.0000,-150.0000
C01384=-5.000,45.800,87.000,0.0000,0.0000,-150.0000
C01385=-10.000,45.800,87.000,0.0000,0.0000,-150.0000
C01386=-15.000,45.800,87.000,0.0000,0.0000,-150.0000
C01387=-20.000,45.800,87.000,0.0000,0.0000,-150.0000
C01388=-25.000,45.800,87.000,0.0000,0.0000,-150.0000
C01389=-30.000,45.800,87.000,0.0000,0.0000,-150.0000
C01390=-35.000,45.800,87.000,0.0000,0.0000,-150.0000
C01391=-40.000,45.800,87.000,0.0000,0.0000,-150.0000
C01392=-45.000,45.800,87.000,0.0000,0.0000,-150.0000
C01393=-50.000,45.800,87.000,0.0000,0.0000,-150.0000
C01394=-55.000,45.800,87.000,0.0000,0.0000,-150.0000
C01395=-60.000,45.800,87.000,0.0000,0.0000,-150.0000
C01396=-65.000,45.800,87.000,0.0000,0.0000,-150.0000
C01397=-70.000,45.800,87.000,0.0000,0.0000,-150.0000
C01398=-75.000,45.800,87.000,0.0000,0.0000,-150.0000
C01399=-76.950,43.850,87.000,0.0000,0.0000,-150.0000
C01400=-75.000,41.900,87.000,0.0000,0.0000,-150.0000
C01401=-70.195,41.900,87.000,0.0000,0.0000,-150.0000
C01402=-65.390,41.900,87.000,0.0000,0.0000,-150.0000
C01403=-60.585,41.900,87.000,0.0000,0.0000,-150.0000
C01404=-55.780,41.900,87.000,0.0000,0.0000,-150.0000
C01405=-50.975,41.900,87.000,0.0000,0.0000,-150.0000
C01406=-46.170,41.900,87.000,0.0000,0.0000,-150.0000
C01407=-41.365,41.900,87.000,0.0000,0.0000,-150.0000
C01408=-36.560,41.900,87.000,0.0000,0.0000,-150.0000
C01409=-31.755,41.900,87.000,0.0000,0.0000,-150.0000
C01410=-26.950,41.900,87.000,0.0000,0.0000,-150.0000
C01411=-26.950,36.900,87.000,0.0000,0.0000,-150.0000
C01412=-26.950,31.900,87.000,0.0000,0.0000,-150.0000
C01413=-26.950,26.900,87.000,0.0000,0.0000,-150.0000
C01414=-26.950,21.900,87.000,0.0000,0.0000,-150.0000
C01415=-26.950,16.900,87.000,0.0000,0.0000,-150.0000
C01416=-26.950,11.900,87.000,0.0000,0.0000,-150.0000
C01417=-26.950,6.900,87.000,0.0000,0.0000,-150.0000
C01418=-26.950,1.900,87.000,0.0000,0.0000,-150.0000
C01419=-26.950,-3.100,87.000,0.0000,0.0000,-150.0000
C01420=-26.950,-8.100,87.000,0.0000,0.0000,-150.0000
C01421=-26.950,-13.100,87.000,0.0000,0.0000,-150.0000
C01422=-26.950,-18.100,87.000,0.0000,0.0000,-150.0000
C01423=-26.950,-23.100,87.000,0.0000,0.0000,-150.0000
C01424=-26.950,-28.100,87.000,0.0000,0.0000,-150.0000
C01425=-26.950,-33.100,87.000,0.0000,0.0000,-150.0000
C01426=-26.950,-38.100,87.000,0.0000,0.0000,-150.0000
C01427=-26.950,-43.100,87.000,0.0000,0.0000,-150.0000
C01428=-26.950,-48.100,87.000,0.0000,0.0000,-150.0000
C01429=-26.950,-53.100,87.000,0.0000,0.0000,-150.0000
C01430=-26.950,-58.100,87.000,0.0000,0.0000,-150.0000
C01431=-26.950,-63.100,87.000,0.0000,0.0000,-150.0000
C01432=-26.950,-68.100,87.000,0.0000,0.0000,-150.0000
C01433=-31.755,-68.100,87.000,0.0000,0.0000,-150.0000
C01434=-36.560,-68.100,87.000,0.0000,0.0000,-150.0000
C01435=-41.365,-68.100,87.000,0.0000,0.0000,-150.0000
C01436=-46.170,-68.100,87.000,0.0000,0.0000,-150.0000
C01437=-50.975,-68.100,87.000,0.0000,0.0000,-150.0000
C01438=-55.780,-68.100,87.000,0.0000,0.0000,-150.0000
C01439=-60.585,-68.100,87.000,0.0000,0.0000,-150.0000
C01440=-65.390,-68.100,87.000,0.0000,0.0000,-150.0000
C01441=-70.195,-68.100,87.000,0.0000,0.0000,-150.0000
C01442=-75.000,-68.100,87.000,0.0000,0.0000,-150.0000
C01443=-75.000,-68.100,88.700,0.0000,0.0000,-150.0000
C01444=-70.195,-68.100,88.700,0.0000,0.0000,-150.0000
C01445=-65.390,-68.100,88.700,0.0000,0.0000,-150.0000
C01446=-60.585,-68.100,88.700,0.0000,0.0000,-150.0000
C01447=-55.780,-68.100,88.700,0.0000,0.0000,-150.0000
C01448=-50.975,-68.100,88.700,0.0000,0.0000,-150.0000
C01449=-46.170,-68.100,88.700,0.0000,0.0000,-150.0000
C01450=-41.365,-68.100,88.700,0.0000,0.0000,-150.0000
C01451=-36.560,-68.100,88.700,0.0000,0.0000,-150.0000
C01452=-31.755,-68.100,88.700,0.0000,0.0000,-150.0000
C01453=-26.950,-68.100,88.700,0.0000,0.0000,-150.0000
C01454=-26.950,-63.100,88.700,0.0000,0.0000,-150.0000
C01455=-26.950,-58.100,88.700,0.0000,0.0000,-150.0000
C01456=-26.950,-53.100,88.700,0.0000,0.0000,-150.0000
C01457=-26.950,-48.100,88.700,0.0000,0.0000,-150.0000
C01458=-26.950,-43.100,88.700,0.0000,0.0000,-150.0000
C01459=-26.950,-38.100,88.700,0.0000,0.0000,-150.0000
C01460=-26.950,-33.100,88.700,0.0000,0.0000,-150.0000
C01461=-26.950,-28.100,88.700,0.0000,0.0000,-150.0000
C01462=-26.950,-23.100,88.700,0.0000,0.0000,-150.0000
C01463=-26.950,-18.100,88.700,0.0000,0.0000,-150.0000
C01464=-26.950,-13.100,88.700,0.0000,0.0000,-150.0000
C01465=-26.950,-8.100,88.700,0.0000,0.0000,-150.0000
C01466=-26.950,-3.100,88.700,0.0000,0.0000,-150.0000
C01467=-26.950,1.900,88.700,0.0000,0.0000,-150.0000
C01468=-26.950,6.900,88.700,0.0000,0.0000,-150.0000
C01469=-26.950,11.900,88.700,0.0000,0.0000,-150.0000
C01470=-26.950,16.900,88.700,0.0000,0.0000,-150.0000
C01471=-26.950,21.900,88.700,0.0000,0.0000,-150.0000
C01472=-26.950,26.900,88.700,0.0000,0.0000,-150.0000
C01473=-26.950,31.900,88.700,0.0000,0.0000,-150.0000
C01474=-26.950,36.900,88.700,0.0000,0.0000,-150.0000
C01475=-26.950,41.900,88.700,0.0000,0.0000,-150.0000
C01476=-31.733,41.900,88.700,0.0000,0.0000,-150.0000
C01477=-36.517,41.900,88.700,0.0000,0.0000,-150.0000
C01478=-41.300,41.900,88.700,0.0000,0.0000,-150.0000
C01479=-46.083,41.900,88.700,0.0000,0.0000,-150.0000
C01480=-50.867,41.900,88.700,0.0000,0.0000,-150.0000
C01481=-55.650,41.900,88.700,0.0000,0.0000,-150.0000
C01482=-60.433,41.900,88.700,0.0000,0.0000,-150.0000
C01483=-65.217,41.900,88.700,0.0000,0.0000,-150.0000
C01484=-70.000,41.900,88.700,0.0000,0.0000,-150.0000
C01485=-75.000,41.900,88.700,0.0000,0.0000,-150.0000
C01486=-76.950,43.850,88.700,0.0000,0.0000,-150.0000
C01487=-75.000,45.800,88.700,0.0000,0.0000,-150.0000
C01488=-70.000,45.800,88.700,0.0000,0.0000,-150.0000
C01489=-65.000,45.800,88.700,0.0000,0.0000,-150.0000
C01490=-60.000,45.800,88.700,0.0000,0.0000,-150.0000
C01491=-55.000,45.800,88.700,0.0000,0.0000,-150.0000
C01492=-50.000,45.800,88.700,0.0000,0.0000,-150.0000
C01493=-45.000,45.800,88.700,0.0000,0.0000,-150.0000
C01494=-40.000,45.800,88.700,0.0000,0.0000,-150.0000
C01495=-35.000,45.800,88.700,0.0000,0.0000,-150.0000
C01496=-30.000,45.800,88.700,0.0000,0.0000,-150.0000
C01497=-25.000,45.800,88.700,0.0000,0.0000,-150.0000
C01498=-20.000,45.800,88.700,0.0000,0.0000,-150.0000
C01499=-15.000,45.800,88.700,0.0000,0.0000,-150.0000
C01500=-10.000,45.800,88.700,0.0000,0.0000,-150.0000
C01501=-5.000,45.800,88.700,0.0000,0.0000,-150.0000
C01502=0.000,45.800,88.700,0.0000,0.0000,-150.0000
C01503=5.000,45.800,88.700,0.0000,0.0000,-150.0000
C01504=10.000,45.800,88.700,0.0000,0.0000,-150.0000
C01505=15.000,45.800,88.700,0.0000,0.0000,-150.0000
C01506=20.000,45.800,88.700,0.0000,0.0000,-150.0000
C01507=25.000,45.800,88.700,0.0000,0.0000,-150.0000
C01508=26.950,43.850,88.700,0.0000,0.0000,-150.0000
C01509=25.000,41.900,88.700,0.0000,0.0000,-150.0000
C01510=20.195,41.900,88.700,0.0000,0.0000,-150.0000
C01511=15.390,41.900,88.700,0.0000,0.0000,-150.0000
C01512=10.585,41.900,88.700,0.0000,0.0000,-150.0000
C01513=5.780,41.900,88.700,0.0000,0.0000,-150.0000
C01514=0.975,41.900,88.700,0.0000,0.0000,-150.0000
C01515=-3.830,41.900,88.700,0.0000,0.0000,-150.0000
C01516=-8.635,41.900,88.700,0.0000,0.0000,-150.0000
C01517=-13.440,41.900,88.700,0.0000,0.0000,-150.0000
C01518=-18.245,41.900,88.700,0.0000,0.0000,-150.0000
C01519=-23.050,41.900,88.700,0.0000,0.0000,-150.0000
C01520=-23.050,36.900,88.700,0.0000,0.0000,-150.0000
C01521=-23.050,31.900,88.700,0.0000,0.0000,-150.0000
C01522=-23.050,26.900,88.700,0.0000,0.0000,-150.0000
C01523=-23.050,21.900,88.700,0.0000,0.0000,-150.0000
C01524=-23.050,16.900,88.700,0.0000,0.0000,-150.0000
C01525=-23.050,11.900,88.700,0.0000,0.0000,-150.0000
C01526=-23.050,6.900,88.700,0.0000,0.0000,-150.0000
C01527=-23.050,1.900,88.700,0.0000,0.0000,-150.0000
C01528=-23.050,-3.100,88.700,0.0000,0.0000,-150.0000
C01529=-23.050,-8.100,88.700,0.0000,0.0000,-150.0000
C01530=-23.050,-13.100,88.700,0.0000,0.0000,-150.0000
C01531=-23.050,-18.100,88.700,0.0000,0.0000,-150.0000
C01532=-23.050,-23.100,88.700,0.0000,0.0000,-150.0000
C01533=-23.050,-28.100,88.700,0.0000,0.0000,-150.0000
C01534=-23.050,-33.100,88.700,0.0000,0.0000,-150.0000
C01535=-23.050,-38.100,88.700,0.0000,0.0000,-150.0000
C01536=-23.050,-43.100,88.700,0.0000,0.0000,-150.0000
C01537=-23.050,-48.100,88.700,0.0000,0.0000,-150.0000
C01538=-23.050,-53.100,88.700,0.0000,0.0000,-150.0000
C01539=-23.050,-58.100,88.700,0.0000,0.0000,-150.0000
C01540=-23.050,-63.100,88.700,0.0000,0.0000,-150.0000
C01541=-23.050,-68.100,88.700,0.0000,0.0000,-150.0000
C01542=-18.267,-68.100,88.700,0.0000,0.0000,-150.0000
C01543=-13.483,-68.100,88.700,0.0000,0.0000,-150.0000
C01544=-8.700,-68.100,88.700,0.0000,0.0000,-150.0000
C01545=-3.917,-68.100,88.700,0.0000,0.0000,-150.0000
C01546=0.867,-68.100,88.700,0.0000,0.0000,-150.0000
C01547=5.650,-68.100,88.700,0.0000,0.0000,-150.0000
C01548=10.433,-68.100,88.700,0.0000,0.0000,-150.0000
C01549=15.217,-68.100,88.700,0.0000,0.0000,-150.0000
C01550=20.000,-68.100,88.700,0.0000,0.0000,-150.0000
C01551=25.000,-68.100,88.700,0.0000,0.0000,-150.0000
C01552=26.950,-70.050,88.700,0.0000,0.0000,-150.0000
C01553=25.000,-72.000,88.700,0.0000,0.0000,-150.0000
C01554=20.000,-72.000,88.700,0.0000,0.0000,-150.0000
C01555=15.000,-72.000,88.700,0.0000,0.0000,-150.0000
C01556=10.000,-72.000,88.700,0.0000,0.0000,-150.0000
C01557=5.000,-72.000,88.700,0.0000,0.0000,-150.0000
C01558=0.000,-72.000,88.700,0.0000,0.0000,-150.0000
C01559=-5.000,-72.000,88.700,0.0000,0.0000,-150.0000
C01560=-10.000,-72.000,88.700,0.0000,0.0000,-150.0000
C01561=-15.000,-72.000,88.700,0.0000,0.0000,-150.0000
C01562=-20.000,-72.000,88.700,0.0000,0.0000,-150.0000
C01563=-25.000,-72.000,88.700,0.0000,0.0000,-150.0000
C01564=-30.000,-72.000,88.700,0.0000,0.0000,-150.0000
C01565=-35.000,-72.000,88.700,0.0000,0.0000,-150.0000
C01566=-40.000,-72.000,88.700,0.0000,0.0000,-150.0000
C01567=-45.000,-72.000,88.700,0.0000,0.0000,-150.0000
C01568=-50.000,-72.000,88.700,0.0000,0.0000,-150.0000
C01569=-55.000,-72.000,88.700,0.0000,0.0000,-150.0000
C01570=-60.000,-72.000,88.700,0.0000,0.0000,-150.0000
C01571=-65.000,-72.000,88.700,0.0000,0.0000,-150.0000
C01572=-70.000,-72.000,88.700,0.0000,0.0000,-150.0000
C01573=-75.000,-72.000,88.700,0.0000,0.0000,-150.0000
C01574=-75.000,-72.000,90.400,0.0000,0.0000,-150.0000
C01575=-70.000,-72.000,90.400,0.0000,0.0000,-150.0000
C01576=-65.000,-72.000,90.400,0.0000,0.0000,-150.0000
C01577=-60.000,-72.000,90.400,0.0000,0.0000,-150.0000
C01578=-55.000,-72.000,90.400,0.0000,0.0000,-150.0000
C01579=-50.000,-72.000,90.400,0.0000,0.0000,-150.0000
C01580=-45.000,-72.000,90.400,0.0000,0.0000,-150.0000
C01581=-40.000,-72.000,90.400,0.0000,0.0000,-150.0000
C01582=-35.000,-72.000,90.400,0.0000,0.0000,-150.0000
C01583=-30.000,-72.000,90.400,0.0000,0.0000,-150.0000
C01584=-25.000,-72.000,90.400,0.0000,0.0000,-150.0000
C01585=-20.000,-72.000,90.400,0.0000,0.0000,-150.0000
C01586=-15.000,-72.000,90.400,0.0000,0.0000,-150.0000
C01587=-10.000,-72.000,90.400,0.0000,0.0000,-150.0000
C01588=-5.000,-72.000,90.400,0.0000,0.0000,-150.0000
C01589=0.000,-72.000,90.400,0.0000,0.0000,-150.0000
C01590=5.000,-72.000,90.400,0.0000,0.0000,-150.0000
C01591=10.000,-72.000,90.400,0.0000,0.0000,-150.0000
C01592=15.000,-72.000,90.400,0.0000,0.0000,-150.0000
C01593=20.000,-72.000,90.400,0.0000,0.0000,-150.0000
C01594=25.000,-72.000,90.400,0.0000,0.0000,-150.0000
C01595=26.950,-70.050,90.400,0.0000,0.0000,-150.0000
C01596=25.000,-68.100,90.400,0.0000,0.0000,-150.0000
C01597=20.195,-68.100,90.400,0.0000,0.0000,-150.0000
C01598=15.390,-68.100,90.400,0.0000,0.0000,-150.0000
C01599=10.585,-68.100,90.400,0.0000,0.0000,-150.0000
C01600=5.780,-68.100,90.400,0.0000,0.0000,-150.0000
C01601=0.975,-68.100,90.400,0.0000,0.0000,-150.0000
C01602=-3.830,-68.100,90.400,0.0000,0.0000,-150.0000
C01603=-8.635,-68.100,90.400,0.0000,0.0000,-150.0000
C01604=-13.440,-68.100,90.400,0.0000,0.0000,-150.0000
C01605=-18.245,-68.100,90.400,0.0000,0.0000,-150.0000
C01606=-23.050,-68.100,90.400,0.0000,0.0000,-150.0000
C01607=-23.050,-63.100,90.400,0.0000,0.0000,-150.0000
C01608=-23.050,-58.100,90.400,0.0000,0.0000,-150.0000
C01609=-23.050,-53.100,90.400,0.0000,0.0000,-150.0000
C01610=-23.050,-48.100,90.400,0.0000,0.0000,-150.0000
C01611=-23.050,-43.100,90.400,0.0000,0.0000,-150.0000
C01612=-23.050,-38.100,90.400,0.0000,0.0000,-150.0000
C01613=-23.050,-33.100,90.400,0.0000,0.0000,-150.0000
C01614=-23.050,-28.100,90.400,0.0000,0.0000,-150.0000
C01615=-23.050,-23.100,90.400,0.0000,0.0000,-150.0000
C01616=-23.050,-18.100,90.400,0.0000,0.0000,-150.0000
C01617=-23.050,-13.100,90.400,0.0000,0.0000,-150.0000
C01618=-23.050,-8.100,90.400,0.0000,0.0000,-150.0000
C01619=-23.050,-3.100,90.400,0.0000,0.0000,-150.0000
C01620=-23.050,1.900,90.400,0.0000,0.0000,-150.0000
C01621=-23.050,6.900,90.400,0.0000,0.0000,-150.0000
C01622=-23.050,11.900,90.400,0.0000,0.0000,-150.0000
C01623=-23.050,16.900,90.400,0.0000,0.0000,-150.0000
C01624=-23.050,21.900,90.400,0.0000,0.0000,-150.0000
C01625=-23.050,26.900,90.400,0.0000,0.0000,-150.0000
C01626=-23.050,31.900,90.400,0.0000,0.0000,-150.0000
C01627=-23.050,36.900,90.400,0.0000,0.0000,-150.0000
C01628=-23.050,41.900,90.400,0.0000,0.0000,-150.0000
C01629=-18.267,41.900,90.400,0.0000,0.0000,-150.0000
C01630=-13.483,41.900,90.400,0.0000,0.0000,-150.0000
C01631=-8.700,41.900,90.400,0.0000,0.0000,-150.0000
C01632=-3.917,41.900,90.400,0.0000,0.0000,-150.0000
C01633=0.867,41.900,90.400,0.0000,0.0000,-150.0000
C01634=5.650,41.900,90.400,0.0000,0.0000,-150.0000
C01635=10.433,41.900,90.400,0.0000,0.0000,-150.0000
C01636=15.217,41.900,90.400,0.0000,0.0000,-150.0000
C01637=20.000,41.900,90.400,0.0000,0.0000,-150.0000
C01638=25.000,41.900,90.400,0.0000,0.0000,-150.0000
C01639=26.950,43.850,90.400,0.0000,0.0000,-150.0000
C01640=25.000,45.800,90.400,0.0000,0.0000,-150.0000
C01641=20.000,45.800,90.400,0.0000,0.0000,-150.0000
C01642=15.000,45.800,90.400,0.0000,0.0000,-150.0000
C01643=10.000,45.800,90.400,0.0000,0.0000,-150.0000
C01644=5.000,45.800,90.400,0.0000,0.0000,-150.0000
C01645=0.000,45.800,90.400,0.0000,0.0000,-150.0000
C01646=-5.000,45.800,90.400,0.0000,0.0000,-150.0000
C01647=-10.000,45.800,90.400,0.0000,0.0000,-150.0000
C01648=-15.000,45.800,90.400,0.0000,0.0000,-150.0000
C01649=-20.000,45.800,90.400,0.0000,0.0000,-150.0000
C01650=-25.000,45.800,90.400,0.0000,0.0000,-150.0000
C01651=-30.000,45.800,90.400,0.0000,0.0000,-150.0000
C01652=-35.000,45.800,90.400,0.0000,0.0000,-150.0000
C01653=-40.000,45.800,90.400,0.0000,0.0000,-150.0000
C01654=-45.000,45.800,90.400,0.0000,0.0000,-150.0000
C01655=-50.000,45.800,90.400,0.0000,0.0000,-150.0000
C01656=-55.000,45.800,90.400,0.0000,0.0000,-150.0000
C01657=-60.000,45.800,90.400,0.0000,0.0000,-150.0000
C01658=-65.000,45.800,90.400,0.0000,0.0000,-150.0000
C01659=-70.000,45.800,90.400,0.0000,0.0000,-150.0000
C01660=-75.000,45.800,90.400,0.0000,0.0000,-150.0000
C01661=-76.950,43.850,90.400,0.0000,0.0000,-150.0000
C01662=-75.000,41.900,90.400,0.0000,0.0000,-150.0000
C01663=-70.195,41.900,90.400,0.0000,0.0000,-150.0000
C01664=-65.390,41.900,90.400,0.0000,0.0000,-150.0000
C01665=-60.585,41.900,90.400,0.0000,0.0000,-150.0000
C01666=-55.780,41.900,90.400,0.0000,0.0000,-150.0000
C01667=-50.975,41.900,90.400,0.0000,0.0000,-150.0000
C01668=-46.170,41.900,90.400,0.0000,0.0000,-150.0000
C01669=-41.365,41.900,90.400,0.0000,0.0000,-150.0000
C01670=-36.560,41.900,90.400,0.0000,0.0000,-150.0000
C01671=-31.755,41.900,90.400,0.0000,0.0000,-150.0000
C01672=-26.950,41.900,90.400,0.0000,0.0000,-150.0000
C01673=-26.950,36.900,90.400,0.0000,0.0000,-150.0000
C01674=-26.950,31.900,90.400,0.0000,0.0000,-150.0000
C01675=-26.950,26.900,90.400,0.0000,0.0000,-150.0000
C01676=-26.950,21.900,90.400,0.0000,0.0000,-150.0000
C01677=-26.950,16.900,90.400,0.0000,0.0000,-150.0000
C01678=-26.950,11.900,90.400,0.0000,0.0000,-150.0000
C01679=-26.950,6.900,90.400,0.0000,0.0000,-150.0000
C01680=-26.950,1.900,90.400,0.0000,0.0000,-150.0000
C01681=-26.950,-3.100,90.400,0.0000,0.0000,-150.0000
C01682=-26.950,-8.100,90.400,0.0000,0.0000,-150.0000
C01683=-26.950,-13.100,90.400,0.0000,0.0000,-150.0000
C01684=-26.950,-18.100,90.400,0.0000,0.0000,-150.0000
C01685=-26.950,-23.100,90.400,0.0000,0.0000,-150.0000
C01686=-26.950,-28.100,90.400,0.0000,0.0000,-150.0000
C01687=-26.950,-33.100,90.400,0.0000,0.0000,-150.0000
C01688=-26.950,-38.100,90.400,0.0000,0.0000,-150.0000
C01689=-26.950,-43.100,90.400,0.0000,0.0000,-150.0000
C01690=-26.950,-48.100,90.400,0.0000,0.0000,-150.0000
C01691=-26.950,-53.100,90.400,0.0000,0.0000,-150.0000
C01692=-26.950,-58.100,90.400,0.0000,0.0000,-150.0000
C01693=-26.950,-63.100,90.400,0.0000,0.0000,-150.0000
C01694=-26.950,-68.100,90.400,0.0000,0.0000,-150.0000
C01695=-31.755,-68.100,90.400,0.0000,0.0000,-150.0000
C01696=-36.560,-68.100,90.400,0.0000,0.0000,-150.0000
C01697=-41.365,-68.100,90.400,0.0000,0.0000,-150.0000
C01698=-46.170,-68.100,90.400,0.0000,0.0000,-150.0000
C01699=-50.975,-68.100,90.400,0.0000,0.0000,-150.0000
C01700=-55.780,-68.100,90.400,0.0000,0.0000,-150.0000
C01701=-60.585,-68.100,90.400,0.0000,0.0000,-150.0000
C01702=-65.390,-68.100,90.400,0.0000,0.0000,-150.0000
C01703=-70.195,-68.100,90.400,0.0000,0.0000,-150.0000
C01704=-75.000,-68.100,90.400,0.0000,0.0000,-150.0000
C01705=-75.000,-68.100,92.100,0.0000,0.0000,-150.0000
C01706=-70.195,-68.100,92.100,0.0000,0.0000,-150.0000
C01707=-65.390,-68.100,92.100,0.0000,0.0000,-150.0000
C01708=-60.585,-68.100,92.100,0.0000,0.0000,-150.0000
C01709=-55.780,-68.100,92.100,0.0000,0.0000,-150.0000
C01710=-50.975,-68.100,92.100,0.0000,0.0000,-150.0000
C01711=-46.170,-68.100,92.100,0.0000,0.0000,-150.0000
C01712=-41.365,-68.100,92.100,0.0000,0.0000,-150.0000
C01713=-36.560,-68.100,92.100,0.0000,0.0000,-150.0000
C01714=-31.755,-68.100,92.100,0.0000,0.0000,-150.0000
C01715=-26.950,-68.100,92.100,0.0000,0.0000,-150.0000
C01716=-26.950,-63.100,92.100,0.0000,0.0000,-150.0000
C01717=-26.950,-58.100,92.100,0.0000,0.0000,-150.0000
C01718=-26.950,-53.100,92.100,0.0000,0.0000,-150.0000
C01719=-26.950,-48.100,92.100,0.0000,0.0000,-150.0000
C01720=-26.950,-43.100,92.100,0.0000,0.0000,-150.0000
C01721=-26.950,-38.100,92.100,0.0000,0.0000,-150.0000
C01722=-26.950,-33.100,92.100,0.0000,0.0000,-150.0000
C01723=-26.950,-28.100,92.100,0.0000,0.0000,-150.0000
C01724=-26.950,-23.100,92.100,0.0000,0.0000,-150.0000
C01725=-26.950,-18.100,92.100,0.0000,0.0000,-150.0000
C01726=-26.950,-13.100,92.100,0.0000,0.0000,-150.0000
C01727=-26.950,-8.100,92.100,0.0000,0.0000,-150.0000
C01728=-26.950,-3.100,92.100,0.0000,0.0000,-150.0000
C01729=-26.950,1.900,92.100,0.0000,0.0000,-150.0000
C01730=-26.950,6.900,92.100,0.0000,0.0000,-150.0000
C01731=-26.950,11.900,92.100,0.0000,0.0000,-150.0000
C01732=-26.950,16.900,92.100,0.0000,0.0000,-150.0000
C01733=-26.950,21.900,92.100,0.0000,0.0000,-150.0000
C01734=-26.950,26.900,92.100,0.0000,0.0000,-150.0000
C01735=-26.950,31.900,92.100,0.0000,0.0000,-150.0000
C01736=-26.950,36.900,92.100,0.0000,0.0000,-150.0000
C01737=-26.950,41.900,92.100,0.0000,0.0000,-150.0000
C01738=-31.733,41.900,92.100,0.0000,0.0000,-150.0000
C01739=-36.517,41.900,92.100,0.0000,0.0000,-150.0000
C01740=-41.300,41.900,92.100,0.0000,0.0000,-150.0000
C01741=-46.083,41.900,92.100,0.0000,0.0000,-150.0000
C01742=-50.867,41.900,92.100,0.0000,0.0000,-150.0000
C01743=-55.650,41.900,92.100,0.0000,0.0000,-150.0000
C01744=-60.433,41.900,92.100,0.0000,0.0000,-150.0000
C01745=-65.217,41.900,92.100,0.0000,0.0000,-150.0000
C01746=-70.000,41.900,92.100,0.0000,0.0000,-150.0000
C01747=-75.000,41.900,92.100,0.0000,0.0000,-150.0000
C01748=-76.950,43.850,92.100,0.0000,0.0000,-150.0000
C01749=-75.000,45.800,92.100,0.0000,0.0000,-150.0000
C01750=-70.000,45.800,92.100,0.0000,0.0000,-150.0000
C01751=-65.000,45.800,92.100,0.0000,0.0000,-150.0000
C01752=-60.000,45.800,92.100,0.0000,0.0000,-150.0000
C01753=-55.000,45.800,92.100,0.0000,0.0000,-150.0000
C01754=-50.000,45.800,92.100,0.0000,0.0000,-150.0000
C01755=-45.000,45.800,92.100,0.0000,0.0000,-150.0000
C01756=-40.000,45.800,92.100,0.0000,0.0000,-150.0000
C01757=-35.000,45.800,92.100,0.0000,0.0000,-150.0000
C01758=-30.000,45.800,92.100,0.0000,0.0000,-150.0000
C01759=-25.000,45.800,92.100,0.0000,0.0000,-150.0000
C01760=-20.000,45.800,92.100,0.0000,0.0000,-150.0000
C01761=-15.000,45.800,92.100,0.0000,0.0000,-150.0000
C01762=-10.000,45.800,92.100,0.0000,0.0000,-150.0000
C01763=-5.000,45.800,92.100,0.0000,0.0000,-150.0000
C01764=0.000,45.800,92.100,0.0000,0.0000,-150.0000
C01765=5.000,45.800,92.100,0.0000,0.0000,-150.0000
C01766=10.000,45.800,92.100,0.0000,0.0000,-150.0000
C01767=15.000,45.800,92.100,0.0000,0.0000,-150.0000
C01768=20.000,45.800,92.100,0.0000,0.0000,-150.0000
C01769=25.000,45.800,92.100,0.0000,0.0000,-150.0000
C01770=26.950,43.850,92.100,0.0000,0.0000,-150.0000
C01771=25.000,41.900,92.100,0.0000,0.0000,-150.0000
C01772=20.195,41.900,92.100,0.0000,0.0000,-150.0000
C01773=15.390,41.900,92.100,0.0000,0.0000,-150.0000
C01774=10.585,41.900,92.100,0.0000,0.0000,-150.0000
C01775=5.780,41.900,92.100,0.0000,0.0000,-150.0000
C01776=0.975,41.900,92.100,0.0000,0.0000,-150.0000
C01777=-3.830,41.900,92.100,0.0000,0.0000,-150.0000
C01778=-8.635,41.900,92.100,0.0000,0.0000,-150.0000
C01779=-13.440,41.900,92.100,0.0000,0.0000,-150.0000
C01780=-18.245,41.900,92.100,0.0000,0.0000,-150.0000
C01781=-23.050,41.900,92.100,0.0000,0.0000,-150.0000
C01782=-23.050,36.900,92.100,0.0000,0.0000,-150.0000
C01783=-23.050,31.900,92.100,0.0000,0.0000,-150.0000
C01784=-23.050,26.900,92.100,0.0000,0.0000,-150.0000
C01785=-23.050,21.900,92.100,0.0000,0.0000,-150.0000
C01786=-23.050,16.900,92.100,0.0000,0.0000,-150.0000
C01787=-23.050,11.900,92.100,0.0000,0.0000,-150.0000
C01788=-23.050,6.900,92.100,0.0000,0.0000,-150.0000
C01789=-23.050,1.900,92.100,0.0000,0.0000,-150.0000
C01790=-23.050,-3.100,92.100,0.0000,0.0000,-150.0000
C01791=-23.050,-8.100,92.100,0.0000,0.0000,-150.0000
C01792=-23.050,-13.100,92.100,0.0000,0.0000,-150.0000
C01793=-23.050,-18.100,92.100,0.0000,0.0000,-150.0000
C01794=-23.050,-23.100,92.100,0.0000,0.0000,-150.0000
C01795=-23.050,-28.100,92.100,0.0000,0.0000,-150.0000
C01796=-23.050,-33.100,92.100,0.0000,0.0000,-150.0000
C01797=-23.050,-38.100,92.100,0.0000,0.0000,-150.0000
C01798=-23.050,-43.100,92.100,0.0000,0.0000,-150.0000
C01799=-23.050,-48.100,92.100,0.0000,0.0000,-150.0000
C01800=-23.050,-53.100,92.100,0.0000,0.0000,-150.0000
C01801=-23.050,-58.100,92.100,0.0000,0.0000,-150.0000
C01802=-23.050,-63.100,92.100,0.0000,0.0000,-150.0000
C01803=-23.050,-68.100,92.100,0.0000,0.0000,-150.0000
C01804=-18.267,-68.100,92.100,0.0000,0.0000,-150.0000
C01805=-13.483,-68.100,92.100,0.0000,0.0000,-150.0000
C01806=-8.700,-68.100,92.100,0.0000,0.0000,-150.0000
C01807=-3.917,-68.100,92.100,0.0000,0.0000,-150.0000
C01808=0.867,-68.100,92.100,0.0000,0.0000,-150.0000
C01809=5.650,-68.100,92.100,0.0000,0.0000,-150.0000
C01810=10.433,-68.100,92.100,0.0000,0.0000,-150.0000
C01811=15.217,-68.100,92.100,0.0000,0.0000,-150.0000
C01812=20.000,-68.100,92.100,0.0000,0.0000,-150.0000
C01813=25.000,-68.100,92.100,0.0000,0.0000,-150.0000
C01814=26.950,-70.050,92.100,0.0000,0.0000,-150.0000
C01815=25.000,-72.000,92.100,0.0000,0.0000,-150.0000
C01816=20.000,-72.000,92.100,0.0000,0.0000,-150.0000
C01817=15.000,-72.000,92.100,0.0000,0.0000,-150.0000
C01818=10.000,-72.000,92.100,0.0000,0.0000,-150.0000
C01819=5.000,-72.000,92.100,0.0000,0.0000,-150.0000
C01820=0.000,-72.000,92.100,0.0000,0.0000,-150.0000
C01821=-5.000,-72.000,92.100,0.0000,0.0000,-150.0000
C01822=-10.000,-72.000,92.100,0.0000,0.0000,-150.0000
C01823=-15.000,-72.000,92.100,0.0000,0.0000,-150.0000
C01824=-20.000,-72.000,92.100,0.0000,0.0000,-150.0000
C01825=-25.000,-72.000,92.100,0.0000,0.0000,-150.0000
C01826=-30.000,-72.000,92.100,0.0000,0.0000,-150.0000
C01827=-35.000,-72.000,92.100,0.0000,0.0000,-150.0000
C01828=-40.000,-72.000,92.100,0.0000,0.0000,-150.0000
C01829=-45.000,-72.000,92.100,0.0000,0.0000,-150.0000
C01830=-50.000,-72.000,92.100,0.0000,0.0000,-150.0000
C01831=-55.000,-72.000,92.100,0.0000,0.0000,-150.0000
C01832=-60.000,-72.000,92.100,0.0000,0.0000,-150.0000
C01833=-65.000,-72.000,92.100,0.0000,0.0000,-150.0000
C01834=-70.000,-72.000,92.100,0.0000,0.0000,-150.0000
C01835=-75.000,-72.000,92.100,0.0000,0.0000,-150.0000
C01836=-75.000,-72.000,93.800,0.0000,0.0000,-150.0000
C01837=-70.000,-72.000,93.800,0.0000,0.0000,-150.0000
C01838=-65.000,-72.000,93.800,0.0000,0.0000,-150.0000
C01839=-60.000,-72.000,93.800,0.0000,0.0000,-150.0000
C01840=-55.000,-72.000,93.800,0.0000,0.0000,-150.0000
C01841=-50.000,-72.000,93.800,0.0000,0.0000,-150.0000
C01842=-45.000,-72.000,93.800,0.0000,0.0000,-150.0000
C01843=-40.000,-72.000,93.800,0.0000,0.0000,-150.0000
C01844=-35.000,-72.000,93.800,0.0000,0.0000,-150.0000
C01845=-30.000,-72.000,93.800,0.0000,0.0000,-150.0000
C01846=-25.000,-72.000,93.800,0.0000,0.0000,-150.0000
C01847=-20.000,-72.000,93.800,0.0000,0.0000,-150.0000
C01848=-15.000,-72.000,93.800,0.0000,0.0000,-150.0000
C01849=-10.000,-72.000,93.800,0.0000,0.0000,-150.0000
C01850=-5.000,-72.000,93.800,0.0000,0.0000,-150.0000
C01851=0.000,-72.000,93.800,0.0000,0.0000,-150.0000
C01852=5.000,-72.000,93.800,0.0000,0.0000,-150.0000
C01853=10.000,-72.000,93.800,0.0000,0.0000,-150.0000
C01854=15.000,-72.000,93.800,0.0000,0.0000,-150.0000
C01855=20.000,-72.000,93.800,0.0000,0.0000,-150.0000
C01856=25.000,-72.000,93.800,0.0000,0.0000,-150.0000
C01857=26.950,-70.050,93.800,0.0000,0.0000,-150.0000
C01858=25.000,-68.100,93.800,0.0000,0.0000,-150.0000
C01859=20.195,-68.100,93.800,0.0000,0.0000,-150.0000
C01860=15.390,-68.100,93.800,0.0000,0.0000,-150.0000
C01861=10.585,-68.100,93.800,0.0000,0.0000,-150.0000
C01862=5.780,-68.100,93.800,0.0000,0.0000,-150.0000
C01863=0.975,-68.100,93.800,0.0000,0.0000,-150.0000
C01864=-3.830,-68.100,93.800,0.0000,0.0000,-150.0000
C01865=-8.635,-68.100,93.800,0.0000,0.0000,-150.0000
C01866=-13.440,-68.100,93.800,0.0000,0.0000,-150.0000
C01867=-18.245,-68.100,93.800,0.0000,0.0000,-150.0000
C01868=-23.050,-68.100,93.800,0.0000,0.0000,-150.0000
C01869=-23.050,-63.100,93.800,0.0000,0.0000,-150.0000
C01870=-23.050,-58.100,93.800,0.0000,0.0000,-150.0000
C01871=-23.050,-53.100,93.800,0.0000,0.0000,-150.0000
C01872=-23.050,-48.100,93.800,0.0000,0.0000,-150.0000
